_attributesSuccess := THIS^.pLogRecord^.attributes.setStringAttribute(
	key:=key,
	value:=value,
	failureReason=>_attributesFailureReason
);
IF NOT _attributesSuccess THEN
	THIS^._failed := TRUE;
	CASE _attributesFailureReason OF
		E_AttributesFailureReason.MEMORY_ALLOCATION_FAILURE:
			THIS^._failureReason := E_LoggerFailureReason.MEMORY_ALLOCATION_FAILURE;
		E_AttributesFailureReason.ATTRIBUTE_COUNT_LIMIT_REACHED:
			THIS^._failureReason := E_LoggerFailureReason.ATTRIBUTE_COUNT_LIMIT_REACHED;
		E_AttributesFailureReason.KV_VALUE_TYPE_UNSUPPORTED:
			THIS^._failureReason := E_LoggerFailureReason.ATTRIBUTE_VALUE_TYPE_UNSUPPORTED;
	ELSE
		THIS^._failureReason := E_LoggerFailureReason.ATTRIBUTE_VALUE_INVALID;
	END_CASE
END_IF
END_METHOD

METHOD setTimestamp: REFERENCE TO FB_Logger
VAR_INPUT
	timestamp: ULINT;
END_VAR
setTimestamp REF= THIS^;

IF THIS^._shouldReturnEarly() THEN
	RETURN;
END_IF

// if everything above worked, assign the value
THIS^.pLogRecord^.timestamp := timestamp;
END_METHOD

(* Sets the record's trace id from raw bytes. Application code uses setTraceContextFromSpan; this setter is for tests and for setTraceContextFromSpan itself. *)
METHOD _setTraceId: REFERENCE TO FB_Logger
VAR_INPUT
	pBytes: POINTER TO BYTE;
	nSize: UDINT;
END_VAR
VAR
	_pDest: POINTER TO FB_TraceId;
	_factoryFailureReason: E_ValueFactoryFailureReason;
END_VAR
_setTraceId REF= THIS^;

IF THIS^._shouldReturnEarly() THEN
	RETURN;
END_IF

// create an instance of FB_TraceId
IF NOT ValueFactory.createTraceId(
	pDest:=_pDest,
	pBytes:=pBytes,
	nSize:=nSize,
	failureReason=>_factoryFailureReason
	) THEN
	THIS^._failed := TRUE;
	CASE _factoryFailureReason OF
		E_ValueFactoryFailureReason.MEMORY_ALLOCATION_FAILURE:
			THIS^._failureReason := E_LoggerFailureReason.MEMORY_ALLOCATION_FAILURE;
		E_ValueFactoryFailureReason.TRACE_ID_BYTES_POINTER_NULL:
			THIS^._failureReason := E_LoggerFailureReason.TRACE_ID_BYTES_POINTER_NULL;
		E_ValueFactoryFailureReason.TRACE_ID_BYTE_COUNT_TOO_SMALL:
			THIS^._failureReason := E_LoggerFailureReason.TRACE_ID_BYTE_COUNT_TOO_SMALL;
	ELSE
		THIS^._failureReason := E_LoggerFailureReason.TRACE_ID_INVALID;
	END_CASE
	RETURN;
END_IF

// assign to the log record
// delete trace id if it's already set.
IF THIS^.pLogRecord^.traceId <> 0 THEN
	THIS^.pLogRecord^.traceId^.delete(pSelf:=THIS^.pLogRecord^.traceId);
END_IF
// transfer ownership of the data
THIS^.pLogRecord^.traceId := _pDest;
_pDest := 0;
END_METHOD

(*
	This method starts the build process with the required log record state.
	Use the fluent setter methods for optional fields.
	
	Example:
	IF NOT logger
		.startLogRecord(severityNumber := E_SeverityNumber.WARN)
		.setBody('process cycle amps warning, motor fault imminent')
		.setTraceContextFromSpan(pSpan)  // a no-op when pSpan is 0
		.setNumberAttribute('motor.amps.min', minAmps)
		.setNumberAttribute('motor.amps.max', maxAmps)
		.setNumberAttribute('motor.amps.avg', avgAmps)
		.emit(failureResult=>failureResult) THEN
		// CASE failureResult OF ...
	END_IF
*)
METHOD startLogRecord: REFERENCE TO FB_Logger
VAR_INPUT
	severityNumber: E_SeverityNumber;
END_VAR
VAR
	_timestamp: ULINT;
END_VAR
VAR CONSTANT
	UNIX_EPOCH_DIFF: ULINT := 116444736000000000;
END_VAR
startLogRecord REF= THIS^;

// do not replace the first failure in an active fluent chain
IF THIS^.pLogRecord <> 0 THEN
	IF NOT THIS^._failed THEN
		THIS^._failed := TRUE;
		THIS^._failureReason := E_LoggerFailureReason.LOG_RECORD_ALREADY_STARTED;
	END_IF
	RETURN;
END_IF

THIS^._failed := FALSE;
THIS^._failureReason := E_LoggerFailureReason.NA;


_timestamp := (F_GetSystemTime() - UNIX_EPOCH_DIFF) * 100;  // NT ticks (100ns) -> unix epoch nanos


// instantiate a log record
IF NOT THIS^._createLogRecord(
	pDest:=THIS^.pLogRecord,
	severityNumber:=severityNumber,
	timestamp:=_timestamp,
	failureReason=>THIS^._failureReason
	) THEN
	THIS^._failed := TRUE;
END_IF
END_METHOD

END_FUNCTION_BLOCK

// ---- OTEL/LOGGING/PROVIDER/FUNCTION_BLOCKS/FB_LoggerProvider.TcPOU
FUNCTION_BLOCK FB_LoggerProvider
VAR
	_resource: REFERENCE TO FB_Resource; // borrowed; the declaring scope owns its lifetime
	_records: FB_LogRecordQueue(TcOtlp_GVL.MAX_LOG_RECORDS_PER_SCAN);
	_head: POINTER TO ST_LinkedListNode;
	_failureReason: E_LoggerProviderFailureReason;
END_VAR
VAR_OUTPUT
	stagedProcessorCount: UDINT;
END_VAR

METHOD _freeProcessors
VAR
	_idx: UDINT;
	_node: POINTER TO ST_LinkedListNode;
END_VAR
FOR _idx := 0 TO TcOtlp_GVL.MAX_LOOP_COUNT DO
	IF THIS^._head = 0 THEN
		EXIT;
	END_IF
	_node := THIS^._head^.nxt;
	__DELETE(THIS^._head);
	THIS^._head := _node;
	// count down per node, so the count never claims nodes that are gone or hides ones that remain
	IF THIS^.stagedProcessorCount > 0 THEN
		THIS^.stagedProcessorCount := THIS^.stagedProcessorCount - 1;
	END_IF
END_FOR
END_METHOD

//FB_Exit must be implemented explicitly. If there is an implementation, then the
//method is called before the controller removes the code of the function block instance
//(implicit call). The return value is not evaluated.
METHOD FB_Exit: BOOL
VAR_INPUT
    bInCopyCode: BOOL;  // TRUE: the exit method is called in order to leave the instance which will be copied afterwards (online change).  
END_VAR
IF NOT bInCopyCode THEN
	THIS^._freeProcessors();
	THIS^._records.free();
END_IF
END_METHOD

//FB_Init is always available implicitly and it is used primarily for initialization.
//The return value is not evaluated. For a specific influence, you can also declare the
//methods explicitly and provide additional code there with the standard initialization
//code. You can evaluate the return value.
METHOD FB_Init: BOOL
VAR_INPUT
    bInitRetains: BOOL; // TRUE: the retain variables are initialized (reset warm / reset cold)
    bInCopyCode: BOOL;  // TRUE: the instance will be copied to the copy code afterward (online change)
	resource: REFERENCE TO FB_Resource;
END_VAR
THIS^._resource REF= resource;
END_METHOD

METHOD onEmit : BOOL
VAR_IN_OUT
	record: POINTER TO FB_LogRecord;
END_VAR
VAR
	_pushFailureReason: E_LogRecordQueueFailureReason;
END_VAR
onEmit := FALSE;

IF record = 0 THEN
	RETURN;
END_IF

IF NOT THIS^._records.push(pValue:=record, failureReason=>_pushFailureReason) THEN
	RETURN;
END_IF

onEmit := TRUE;
END_METHOD

PROPERTY resource : REFERENCE TO FB_Resource
GET
resource REF= THIS^._resource;
END_GET
END_PROPERTY

METHOD stageProcessor : REFERENCE TO FB_LoggerProvider
VAR_INPUT
	processor: REFERENCE TO FB_LogRecordProcessor_Base;
END_VAR
VAR
	_idx: UDINT;
	_node: POINTER TO ST_LinkedListNode;
END_VAR
stageProcessor REF= THIS^;

// special case if no processors have been registered
IF THIS^._head = 0 THEN
	THIS^._head := __NEW(ST_LinkedListNode);
	IF THIS^._head = 0 THEN
		THIS^._failureReason := E_LoggerProviderFailureReason.STAGE_PROCESSOR_FAILURE;
		RETURN;
	END_IF
	THIS^._head^.val := processor.pSelf;
	THIS^.stagedProcessorCount := THIS^.stagedProcessorCount + 1;
// generic case if at least on processor has been registerd
ELSE
	_node := THIS^._head;
	FOR _idx := 0 TO TcOtlp_GVL.MAX_LOOP_COUNT DO
		IF _node^.val = processor.pSelf THEN
			// silently do nothing if processor already added for this tick
			RETURN;
		ELSIF _node^.nxt = 0 THEN
			// at most MAX_LOOP_COUNT nodes, so _freeProcessors always releases them all
			IF THIS^.stagedProcessorCount >= TcOtlp_GVL.MAX_LOOP_COUNT THEN
				THIS^._failureReason := E_LoggerProviderFailureReason.STAGE_PROCESSOR_FAILURE;
				RETURN;
			END_IF
			_node^.nxt := __NEW(ST_LinkedListNode);
			IF _node^.nxt = 0 THEN
				THIS^._failureReason := E_LoggerProviderFailureReason.STAGE_PROCESSOR_FAILURE;
				RETURN;
			END_IF
			_node^.nxt^.val := processor.pSelf;
			THIS^.stagedProcessorCount := THIS^.stagedProcessorCount + 1;
			RETURN;
		END_IF
		_node := _node^.nxt;
	END_FOR
END_IF
END_METHOD

METHOD tick : BOOL
VAR_OUTPUT
	failureReason: E_LoggerProviderFailureReason;
END_VAR
VAR
	_i: UDINT;
	_j: UDINT;
	_ownedRecordCount: UDINT;
	_node: POINTER TO ST_LinkedListNode;
	_processor: POINTER TO FB_LogRecordProcessor_Base;
	_record: POINTER TO FB_LogRecord;
END_VAR
tick := FALSE;
failureReason := THIS^._failureReason;

// short circuit if fluent calls to add processors failed
IF failureReason <> E_LoggerProviderFailureReason.NA THEN
	RETURN;
END_IF

// if no processors added skip loop iteration and just free the queue
IF THIS^._head = 0 THEN
	THIS^._records.free();
	tick := TRUE;
	RETURN;
END_IF

// loop over each item and call each processor for each record
_ownedRecordCount := THIS^._records.count;
FOR _i := 1 TO _ownedRecordCount DO
	IF NOT THIS^._records.pop(_record) THEN
		failureReason := E_LoggerProviderFailureReason.QUEUE_POP_FAILURE;
		JMP _endLabel;
	END_IF
	// call on emit for each record
	_node := THIS^._head;
	FOR _j := 1 TO THIS^.stagedProcessorCount DO
		IF _node = 0 THEN
			failureReason := E_LoggerProviderFailureReason.UNEXPECTED_NULL_LINKED_LIST_NODE;
			JMP _endLabel;
		END_IF
		_processor := _node^.val;
		IF _processor = 0 THEN
			failureReason := E_LoggerProviderFailureReason.UNEXPECTED_NULL_PROCESSOR_POINTER;
			JMP _endLabel;
		END_IF
		_processor^.onEmit(_record^);
		_node := _node^.nxt;
	END_FOR
	_record^.delete(pSelf:=_record);
END_FOR

// tick each processor
_node := THIS^._head;
FOR _j := 1 TO THIS^.stagedProcessorCount DO
	// guard before dereferencing; walking off the tail on the last iteration is
	// normal termination, so only a list shorter than the count is a failure
	IF _node = 0 THEN
		failureReason := E_LoggerProviderFailureReason.UNEXPECTED_NULL_LINKED_LIST_NODE;
		JMP _endLabel;
	END_IF
	_processor := _node^.val;
	IF _processor = 0 THEN
		failureReason := E_LoggerProviderFailureReason.UNEXPECTED_NULL_PROCESSOR_POINTER;
		JMP _endLabel;
	END_IF
	_processor^.tick();
	_node := _node^.nxt;
END_FOR

// clean up and return
_endLabel:
THIS^._records.free();
THIS^._freeProcessors();
IF _record <> 0 THEN _record^.delete(pSelf:=_record); END_IF
tick := failureReason = E_LoggerProviderFailureReason.NA;
END_METHOD

END_FUNCTION_BLOCK

// ---- OTEL/LOGGING/PROCESSORS/FUNCTION_BLOCKS/FB_LogRecordProcessor_Base.TcPOU
FUNCTION_BLOCK ABSTRACT FB_LogRecordProcessor_Base

METHOD ABSTRACT enrich
VAR_IN_OUT
	logRecord: FB_LogRecord;
END_VAR
END_METHOD

METHOD ABSTRACT free
VAR_INPUT
END_VAR
END_METHOD

METHOD ABSTRACT onEmit
VAR_INPUT
	logRecord: REFERENCE TO FB_LogRecord;
END_VAR
END_METHOD

PROPERTY pSelf : POINTER TO FB_LogRecordProcessor_Base
GET
pSelf := THIS;
END_GET
END_PROPERTY

METHOD ABSTRACT tick
END_METHOD

END_FUNCTION_BLOCK

// ---- OTEL/LOGGING/PROCESSORS/FUNCTION_BLOCKS/FB_LogRecordProcessor_Batch.TcPOU
(*
	Batch processor. onEmit enriches and stores records only. Call the FB body
	cyclically to advance the exporter and export the oldest queued records when
	the schedule delay elapses or a full batch is available.
*)
FUNCTION_BLOCK FB_LogRecordProcessor_Batch EXTENDS FB_LogRecordProcessor_Base;
VAR_OUTPUT
	scheduledDelayMillis: UDINT := 1000;	// maximum delay before queued records are exported
	maxExportBatchSize: UDINT := 512;		// maximum records transferred to one export
	lastOperationSucceeded: BOOL := TRUE;
	failureResult: E_LogRecordProcessorFailureReason;
END_VAR
VAR
	_scheduleDelayTimer: TON;
	_records: FB_LogRecordQueue(maxCount:=0);  // set again during THIS^.FB_Init
	_exporter: REFERENCE TO FB_LogRecordExporter_Base;
	_rejectedCount: UDINT;  // records that could not be cloned or queued
END_VAR

// no-op; override to change log mutation/enrichment functionality
METHOD enrich
VAR_IN_OUT
	logRecord: FB_LogRecord;
END_VAR
END_METHOD

METHOD exportIfNeeded
VAR
	_exportFailureReason: E_LogRecordExporterFailureReason;
END_VAR
IF THIS^.maxExportBatchSize = 0
	OR_ELSE NOT __ISVALIDREF(THIS^._exporter)
	OR_ELSE THIS^._exporter.isBusy()
	OR_ELSE THIS^._records.count = 0 THEN
	RETURN;
END_IF

IF NOT THIS^._scheduleDelayTimer.Q
	AND_THEN THIS^._records.count < THIS^.maxExportBatchSize THEN
	RETURN;
END_IF

IF THIS^._exporter.export(
	logRecords:=THIS^._records,
	count:=THIS^.maxExportBatchSize,
	failureReason=>_exportFailureReason
) THEN
	THIS^._scheduleDelayTimer(IN:=FALSE, PT:=UDINT_TO_TIME(THIS^.scheduledDelayMillis));
	THIS^.lastOperationSucceeded := TRUE;
	THIS^.failureResult := E_LogRecordProcessorFailureReason.NA;
ELSE
	THIS^.lastOperationSucceeded := FALSE;
	THIS^.failureResult := E_LogRecordProcessorFailureReason.EXPORT_FAILURE;
END_IF
END_METHOD

METHOD FB_Exit : BOOL
VAR_INPUT
	bInCopyCode: BOOL;
END_VAR
IF NOT bInCopyCode THEN
	THIS^.free();
END_IF
END_METHOD

//FB_Init is always available implicitly and it is used primarily for initialization.
//The return value is not evaluated. For a specific influence, you can also declare the
//methods explicitly and provide additional code there with the standard initialization
//code. You can evaluate the return value.
METHOD FB_Init: BOOL
VAR_INPUT
    bInitRetains: BOOL; // TRUE: the retain variables are initialized (reset warm / reset cold)
    bInCopyCode: BOOL;  // TRUE: the instance will be copied to the copy code afterward (online change)
	maxQueueSize: UDINT := 2048;			// zero is unbounded; otherwise the oldest record is dropped when full
	scheduledDelayMillis: UDINT := 1000;	// maximum delay before queued records are exported
	maxExportBatchSize: UDINT := 512;		// maximum records transferred to one export
	exporter: REFERENCE TO FB_LogRecordExporter_Base;	// the exporter where the LogRecords are pushed.
END_VAR
THIS^._records.FB_Init(FALSE, FALSE, maxQueueSize);
THIS^.scheduledDelayMillis := scheduledDelayMillis;
THIS^.maxExportBatchSize := maxExportBatchSize;
IF __ISVALIDREF(exporter) THEN
	THIS^._exporter REF= exporter;
END_IF
END_METHOD

METHOD free
THIS^._records.free();
THIS^._scheduleDelayTimer(IN:=FALSE, PT:=UDINT_TO_TIME(THIS^.scheduledDelayMillis));
END_METHOD

(*
	Clones the log record onto the tail of the arrival-order queue.
	When the queue holds maxQueueSize records, the oldest record is
	dropped from the head to make room for the newest.
*)
METHOD onEmit
VAR_INPUT
	logRecord: REFERENCE TO FB_LogRecord;
END_VAR
VAR
	_pRecord: POINTER TO FB_LogRecord;
	_cloneFailureResult: E_LogRecordCloneFailureReason;
	_queueFailureReason: E_LogRecordQueueFailureReason;
END_VAR
THIS^.enrich(logRecord);

IF __ISVALIDREF(THIS^._exporter) THEN
	_pRecord := 0;
	IF NOT logRecord.cloneTo(pDest:=_pRecord, failureReason=>_cloneFailureResult) THEN
		IF _pRecord <> 0 THEN _pRecord^.delete(pSelf:=_pRecord); END_IF
		THIS^._rejectedCount := THIS^._rejectedCount + 1;
		THIS^.lastOperationSucceeded := FALSE;
		THIS^.failureResult := E_LogRecordProcessorFailureReason.RECORD_CLONE_FAILURE;
		RETURN;
	END_IF
	
	IF NOT THIS^._records.push(pValue:=_pRecord, failureReason=>_queueFailureReason) THEN
		_pRecord^.delete(pSelf:=_pRecord);
		THIS^._rejectedCount := THIS^._rejectedCount + 1;
		THIS^.lastOperationSucceeded := FALSE;
		THIS^.failureResult := E_LogRecordProcessorFailureReason.QUEUE_PUSH_FAILURE;
		RETURN;
	END_IF
END_IF

THIS^.lastOperationSucceeded := TRUE;
THIS^.failureResult := E_LogRecordProcessorFailureReason.NA;
END_METHOD

METHOD tick
VAR
	_exportFailureReason: E_LogRecordExporterFailureReason;
END_VAR
THIS^._scheduleDelayTimer(
	IN:=THIS^._records.count > 0,
	PT:=UDINT_TO_TIME(THIS^.scheduledDelayMillis)
);

IF __ISVALIDREF(THIS^._exporter) THEN
	THIS^._exporter.tick(failureReason=>_exportFailureReason);
	THIS^.exportIfNeeded();
END_IF
END_METHOD

(* Records lost so far: evicted from a full queue, or not cloned or queued. *)
PROPERTY droppedCount : UDINT
GET
droppedCount := THIS^._records.droppedCount + THIS^._rejectedCount;
END_GET
END_PROPERTY

(* Records waiting for export. *)
PROPERTY queuedCount : UDINT
GET
queuedCount := THIS^._records.count;
END_GET
END_PROPERTY

END_FUNCTION_BLOCK

// ---- OTEL/LOGGING/PROCESSORS/FUNCTION_BLOCKS/FB_LogRecordProcessor_Simple.TcPOU
FUNCTION_BLOCK FB_LogRecordProcessor_Simple EXTENDS FB_LogRecordProcessor_Base;
VAR
	_records: FB_LogRecordQueue(maxCount:=1);
	_exporter: REFERENCE TO FB_LogRecordExporter_Base;
END_VAR

// no-op, overwride to change log mutation/enrichment functionality
METHOD enrich
VAR_IN_OUT
	logRecord	: FB_LogRecord;
END_VAR
END_METHOD

//FB_Exit must be implemented explicitly. If there is an implementation, then the
//method is called before the controller removes the code of the function block instance
//(implicit call). The return value is not evaluated.
METHOD FB_Exit: BOOL
VAR_INPUT
    bInCopyCode: BOOL;  // TRUE: the exit method is called in order to leave the instance which will be copied afterwards (online change).  
END_VAR
IF NOT bInCopyCode THEN
	THIS^.free();
END_IF
END_METHOD

//FB_Init is always available implicitly and it is used primarily for initialization.
//The return value is not evaluated. For a specific influence, you can also declare the
//methods explicitly and provide additional code there with the standard initialization
//code. You can evaluate the return value.
METHOD FB_Init: BOOL
VAR_INPUT
    bInitRetains: BOOL; // TRUE: the retain variables are initialized (reset warm / reset cold)
    bInCopyCode: BOOL;  // TRUE: the instance will be copied to the copy code afterward (online change)
	exporter: REFERENCE TO FB_LogRecordExporter_Base;
END_VAR
IF __ISVALIDREF(exporter) THEN
	THIS^._exporter REF= exporter;
ELSE
	THIS^._exporter REF= 0;
END_IF
END_METHOD

METHOD free
THIS^._records.free();
END_METHOD

METHOD onEmit
VAR_INPUT
	logRecord: REFERENCE TO FB_LogRecord;
END_VAR
VAR
	_pLogRecord: POINTER TO FB_LogRecord;
	_cloneFailureResult: E_LogRecordCloneFailureReason;
	_queueFailureReason: E_LogRecordQueueFailureReason;
	_exportFailureReason: E_LogRecordExporterFailureReason;
END_VAR
THIS^.enrich(logRecord);

IF __ISVALIDREF(THIS^._exporter) THEN
	IF (NOT THIS^._exporter.isBusy()) THEN
		IF logRecord.cloneTo(pDest:=_pLogRecord, failureReason=>_cloneFailureResult) THEN
			IF THIS^._records.push(pValue:=_pLogRecord, failureReason=>_queueFailureReason) THEN
				THIS^._exporter.export(
					logRecords:=THIS^._records,
					count:=1,
					failureReason=>_exportFailureReason
				);
			END_IF
		END_IF
	END_IF
END_IF

// If the exporter did not accept the buffer, the simple processor drops it.
THIS^.free();
IF _pLogRecord <> 0 THEN _pLogRecord^.delete(pSelf:=_pLogRecord); END_IF
END_METHOD

METHOD tick
VAR
	_exportFailureReason: E_LogRecordExporterFailureReason;
END_VAR
IF __ISVALIDREF(THIS^._exporter) THEN
	THIS^._exporter.tick(failureReason=>_exportFailureReason);
END_IF
END_METHOD

END_FUNCTION_BLOCK

// ---- OTEL/TRACING/EXPORTING/FUNCTION_BLOCKS/FB_SpanExporter_Base.TcPOU
(*
	Contract shared by span exporters. A processor offers a batch with export, which moves up to
	count of the oldest spans out of the processor's queue into the exporter without cloning
	them. The exporter owns the batch until free, which runs when the batch is delivered or
	failed, when the next batch is accepted, and when the exporter is destroyed.
	Concrete exporters advance delivery in tick and report through isBusy whether they can take
	another batch. Only ended spans reach an exporter.
*)
FUNCTION_BLOCK ABSTRACT FB_SpanExporter_Base
VAR
	_spans: FB_SpanQueue(maxCount:=0);
	_exportActive: BOOL;
	_callFailureReason: E_SpanExporterFailureReason;
END_VAR

(*
	Takes ownership of up to count of the oldest spans in spans. While busy it refuses with
	ACTIVE_EXPORT_IN_PROGRESS and leaves spans unchanged. A count of zero accepts nothing and
	succeeds.
*)
METHOD export : BOOL
VAR_IN_OUT
	spans: FB_SpanQueue;  // accepted spans are transferred out of this queue
END_VAR
VAR_INPUT
	count: UDINT;
END_VAR
VAR_OUTPUT
	failureReason: E_SpanExporterFailureReason;
END_VAR
VAR
	_queueFailureReason: E_SpanQueueFailureReason;
END_VAR
export := FALSE;
failureReason := E_SpanExporterFailureReason.NA;

IF THIS^.isBusy() THEN
	failureReason := E_SpanExporterFailureReason.ACTIVE_EXPORT_IN_PROGRESS;
	RETURN;
END_IF

// release a finished batch still held by the exporter before accepting the next one
THIS^.free();
IF NOT spans.transferTo(
	destination:=THIS^._spans,
	count:=count,
	failureReason=>_queueFailureReason
) THEN
	failureReason := E_SpanExporterFailureReason.QUEUE_TRANSFER_FAILURE;
	RETURN;
END_IF

THIS^._exportActive := THIS^._spans.count > 0;
export := TRUE;
END_METHOD

METHOD FB_Exit : BOOL
VAR_INPUT
	bInCopyCode: BOOL;
END_VAR
IF NOT bInCopyCode THEN
	THIS^.free();
END_IF
END_METHOD

(* Releases every span the exporter owns and clears the active export. *)
METHOD free
THIS^._spans.free();
THIS^._exportActive := FALSE;
END_METHOD

(* TRUE while the exporter cannot accept another batch. *)
METHOD ABSTRACT isBusy : BOOL
END_METHOD

(* Advances delivery of the accepted batch. Call it every scan. *)
METHOD ABSTRACT tick : BOOL
VAR_OUTPUT
	failureReason: E_SpanExporterFailureReason;
END_VAR
END_METHOD

END_FUNCTION_BLOCK

// ---- OTEL/TRACING/SPAN/FUNCTION_BLOCKS/FB_SpanQueue.TcPOU
(*
	FIFO queue that owns every FB_Span pointer it contains. push takes ownership and
	clears the caller's pointer; pop hands ownership back. push drops the oldest owned
	spans when the bound is reached. The bound is maxCount, but never more than
	TcOtlp_GVL.MAX_LOOP_COUNT: a maxCount of zero, or one above that limit, is held to
	MAX_LOOP_COUNT so that free always reaches the end.
	reset and next walk the spans oldest first without taking ownership. rotate moves the
	oldest span to the back, so a consumer can skip it and keep arrival order. transferTo moves the oldest spans into another queue, for handing
	a batch to an exporter.
*)
FUNCTION_BLOCK FB_SpanQueue
VAR
	_head: POINTER TO ST_LinkedListNode;
	_tail: POINTER TO ST_LinkedListNode;
	_cursor: POINTER TO ST_LinkedListNode;  // next node returned by next; 0 at the end
END_VAR
VAR_OUTPUT
	count: UDINT;
	maxCount: UDINT;
	droppedCount: UDINT;
END_VAR

(* The enforced bound: maxCount, held to MAX_LOOP_COUNT when it is zero or larger. *)
METHOD _capacity : UDINT
IF THIS^.maxCount = 0 OR THIS^.maxCount > TcOtlp_GVL.MAX_LOOP_COUNT THEN
	_capacity := TcOtlp_GVL.MAX_LOOP_COUNT;
ELSE
	_capacity := THIS^.maxCount;
END_IF
END_METHOD

METHOD FB_Exit : BOOL
VAR_INPUT
	bInCopyCode: BOOL;
END_VAR
IF NOT bInCopyCode THEN
	THIS^.free();
END_IF
END_METHOD

METHOD FB_Init : BOOL
VAR_INPUT
	bInitRetains: BOOL;
	bInCopyCode: BOOL;
	maxCount: UDINT := 0;
END_VAR
THIS^.maxCount := maxCount;
END_METHOD

(*
	Releases every owned span. push holds count to MAX_LOOP_COUNT, so the loop always
	reaches the end. If it ever stops early, the unreleased nodes stay in the queue and
	free returns FALSE, so a later call can finish the job.
*)
METHOD free : BOOL
VAR
	_idx: UDINT;
	_node: POINTER TO ST_LinkedListNode;
	_span: POINTER TO FB_Span;
END_VAR
FOR _idx := 0 TO TcOtlp_GVL.MAX_LOOP_COUNT DO
	IF THIS^._head = 0 THEN
		EXIT;
	END_IF

	_node := THIS^._head;
	THIS^._head := _node^.nxt;
	IF _node^.val <> 0 THEN
		_span := _node^.val;
		_node^.val := 0;
		_span^.delete(pSelf:=_span);
	END_IF
	__DELETE(_node);
	_node := 0;
	IF THIS^.count > 0 THEN
		THIS^.count := THIS^.count - 1;
	END_IF
END_FOR

IF THIS^._head = 0 THEN
	THIS^._tail := 0;
	THIS^.count := 0;
END_IF
THIS^._cursor := THIS^._head;
free := THIS^._head = 0;
END_METHOD

(*
	Returns the span at the cursor and advances it, or 0 after the last span. The span is
	borrowed: the queue still owns it, and it is valid only until it is popped or dropped.
	Call reset first.
*)
METHOD next : POINTER TO FB_Span
next := 0;
IF THIS^._cursor <> 0 THEN
	next := THIS^._cursor^.val;
	THIS^._cursor := THIS^._cursor^.nxt;
END_IF
END_METHOD

(* Moves the oldest span to pValue, which must be 0. The caller owns it on success. *)
METHOD pop : BOOL
VAR_IN_OUT
	pValue: POINTER TO FB_Span;
END_VAR
VAR_OUTPUT
	failureReason: E_SpanQueueFailureReason;
END_VAR
VAR
	_node: POINTER TO ST_LinkedListNode;
END_VAR
pop := FALSE;
failureReason := E_SpanQueueFailureReason.NA;

IF pValue <> 0 THEN
	failureReason := E_SpanQueueFailureReason.DESTINATION_ALREADY_ASSIGNED;
	RETURN;
END_IF
IF THIS^._head = 0 THEN
	failureReason := E_SpanQueueFailureReason.QUEUE_EMPTY;
	RETURN;
END_IF

_node := THIS^._head;
THIS^._head := _node^.nxt;
IF THIS^._head = 0 THEN
	THIS^._tail := 0;
END_IF
IF THIS^._cursor = _node THEN
	THIS^._cursor := THIS^._head;
END_IF

pValue := _node^.val;
_node^.val := 0;
_node^.nxt := 0;
__DELETE(_node);
_node := 0;
THIS^.count := THIS^.count - 1;
pop := failureReason = E_SpanQueueFailureReason.NA;
END_METHOD

(*
	Takes ownership of the span and clears pValue. On failure pValue is left unchanged
	and still owned by the caller.
*)
METHOD push : BOOL
VAR_IN_OUT
	pValue: POINTER TO FB_Span;
END_VAR
VAR_OUTPUT
	failureReason: E_SpanQueueFailureReason;
END_VAR
VAR
	_node: POINTER TO ST_LinkedListNode;
	_droppedSpan: POINTER TO FB_Span;
	_popFailureReason: E_SpanQueueFailureReason;
	_idx: UDINT;
	_bound: UDINT;
END_VAR
push := FALSE;
failureReason := E_SpanQueueFailureReason.NA;

IF pValue = 0 THEN
	failureReason := E_SpanQueueFailureReason.SPAN_POINTER_NULL;
	RETURN;
END_IF

// Allocate before evicting so an allocation failure leaves the queue unchanged.
_node := __NEW(ST_LinkedListNode);
IF _node = 0 THEN
	failureReason := E_SpanQueueFailureReason.MEMORY_ALLOCATION_FAILURE;
	RETURN;
END_IF

// maxCount is writable, so also restore the bound after a runtime reduction.
_bound := THIS^._capacity();
FOR _idx := 0 TO TcOtlp_GVL.MAX_LOOP_COUNT DO
	IF THIS^.count < _bound THEN
		EXIT;
	END_IF
	IF NOT THIS^.pop(pValue:=_droppedSpan, failureReason=>_popFailureReason) THEN
		__DELETE(_node);
		_node := 0;
		failureReason := _popFailureReason;
		RETURN;
	END_IF
	_droppedSpan^.delete(pSelf:=_droppedSpan);
	THIS^.droppedCount := THIS^.droppedCount + 1;
END_FOR
IF THIS^.count >= _bound THEN
	__DELETE(_node);
	_node := 0;
	failureReason := E_SpanQueueFailureReason.MAX_SIZE_ENFORCEMENT_FAILURE;
	RETURN;
END_IF

_node^.val := pValue;
_node^.nxt := 0;
IF THIS^._tail = 0 THEN
	THIS^._head := _node;
ELSE
	THIS^._tail^.nxt := _node;
END_IF
THIS^._tail := _node;
THIS^.count := THIS^.count + 1;
pValue := 0;
push := failureReason = E_SpanQueueFailureReason.NA;
END_METHOD

(* Moves the cursor to the oldest span, so next starts from the head. *)
METHOD reset
THIS^._cursor := THIS^._head;
END_METHOD

(*
	Moves up to count of the oldest spans into destination, which must be empty. Ownership moves
	with the nodes, so nothing is cloned or released. The move stops at this queue's count and at
	the destination's bound.
*)
METHOD transferTo : BOOL
VAR_IN_OUT
	destination: FB_SpanQueue;
END_VAR
VAR_INPUT
	count: UDINT;
END_VAR
VAR_OUTPUT
	failureReason: E_SpanQueueFailureReason;
END_VAR
VAR
	_transferCount: UDINT;
	_idx: UDINT;
END_VAR
transferTo := FALSE;
failureReason := E_SpanQueueFailureReason.NA;

IF ADR(destination) = THIS THEN
	failureReason := E_SpanQueueFailureReason.SELF_TRANSFER_NOT_ALLOWED;
	RETURN;
END_IF
IF destination.count <> 0 OR_ELSE destination._head <> 0 OR_ELSE destination._tail <> 0 THEN
	failureReason := E_SpanQueueFailureReason.DESTINATION_NOT_EMPTY;
	RETURN;
END_IF

_transferCount := MIN(count, THIS^.count, destination._capacity());
IF _transferCount = 0 THEN
	transferTo := TRUE;
	RETURN;
END_IF

// count never exceeds MAX_LOOP_COUNT, so this walk is bounded
destination._head := THIS^._head;
destination._tail := destination._head;
FOR _idx := 1 TO _transferCount - 1 DO
	destination._tail := destination._tail^.nxt;
END_FOR

THIS^._head := destination._tail^.nxt;
destination._tail^.nxt := 0;
destination._cursor := destination._head;
destination.count := _transferCount;

THIS^.count := THIS^.count - _transferCount;
THIS^._cursor := THIS^._head;
IF THIS^._head = 0 THEN
	THIS^._tail := 0;
END_IF
transferTo := TRUE;
END_METHOD

(* Moves the oldest span to the back without changing ownership, and resets the cursor. *)
METHOD rotate : BOOL
VAR_OUTPUT
	failureReason: E_SpanQueueFailureReason;
END_VAR
VAR
	_node: POINTER TO ST_LinkedListNode;
END_VAR
rotate := FALSE;
failureReason := E_SpanQueueFailureReason.NA;

IF THIS^._head = 0 THEN
	failureReason := E_SpanQueueFailureReason.QUEUE_EMPTY;
	RETURN;
END_IF

IF THIS^._head <> THIS^._tail THEN
	_node := THIS^._head;
	THIS^._head := _node^.nxt;
	_node^.nxt := 0;
	THIS^._tail^.nxt := _node;
	THIS^._tail := _node;
END_IF

THIS^._cursor := THIS^._head;
rotate := failureReason = E_SpanQueueFailureReason.NA;
END_METHOD

END_FUNCTION_BLOCK

// ---- OTEL/TRACING/EXPORTING/FUNCTION_BLOCKS/FB_SpanExporter_File.TcPOU
(*
	Appends each accepted batch to a file as one OTLP ProtoJSON TracesData object per line
	(JSON Lines), grouped by resource and scope. The file is opened in append mode and closed
	again for every batch. Call the instance, or tick, every scan: the exporter is busy from
	export until currentState reaches done or error. The batch is released at either end, and
	an error is reported by tick until the next batch is accepted.
*)
FUNCTION_BLOCK FB_SpanExporter_File EXTENDS FB_SpanExporter_Base
VAR_OUTPUT
	currentState: E_FileExporterState;
END_VAR
VAR
	_execute: BOOL;
	_filepath: T_MaxString;
	_hFile: UINT;
	_len: UDINT;
	_execRTrig: R_TRIG;
	_pString: POINTER TO STRING;  // payload buffer, owned while a write is in flight
	_jsonVal: SJsonValue;
	_resourceSpansArray: SJsonValue;
	_fileOpener: FB_FileOpen;
	_fileWriter: FB_FileWrite;
	_fileCloser: FB_FileClose;
	_computedState: E_FileExporterState;
	_failureReason: E_SpanExporterFailureReason;
	_serializationFailureReason: E_ProtoJsonSerializerFailureReason;
	_serializer: FB_SpanProtoJsonSerializer;
END_VAR

THIS^.tick(failureReason=>THIS^._callFailureReason);

METHOD export : BOOL
VAR_IN_OUT
	spans: FB_SpanQueue;
END_VAR
VAR_INPUT
	count: UDINT;
END_VAR
VAR_OUTPUT
	failureReason: E_SpanExporterFailureReason;
END_VAR
// a finished exporter accepts the next batch at once
IF THIS^.currentState = E_FileExporterState.done OR THIS^.currentState = E_FileExporterState.error THEN
	THIS^.currentState := E_FileExporterState.idle;
	THIS^._computedState := E_FileExporterState.idle;
END_IF
export := SUPER^.export(
	spans:=spans,
	count:=count,
	failureReason=>failureReason
);
IF export THEN
	THIS^._failureReason := E_SpanExporterFailureReason.NA;
	THIS^._serializationFailureReason := E_ProtoJsonSerializerFailureReason.NA;
END_IF
END_METHOD

(*
	Releases a payload buffer that is still in flight. The FB_FileWrite reading it is
	destroyed with this instance, so nothing uses the buffer afterwards. TwinCAT then
	runs FB_SpanExporter_Base.FB_Exit, which releases the accepted spans.
*)
METHOD FB_Exit : BOOL
VAR_INPUT
	bInCopyCode: BOOL;  // TRUE: the instance is being copied during an online change
END_VAR
// during an online change the copy keeps the buffer, so it must not be released here
IF NOT bInCopyCode AND _pString <> 0 THEN
	__DELETE(_pString);
	_pString := 0;
END_IF
END_METHOD

METHOD FB_Init : BOOL
VAR_INPUT
	bInitRetains: BOOL;  // TRUE: the retain variables are initialized (reset warm / reset cold)
	bInCopyCode: BOOL;  // TRUE: the instance will be copied to the copy code afterward (online change)
	filepath: T_MaxString;  // file the batches are appended to
END_VAR
THIS^._filepath := filepath;
END_METHOD

METHOD isBusy : BOOL
isBusy := THIS^._exportActive;
END_METHOD

METHOD tick : BOOL
VAR_OUTPUT
	failureReason: E_SpanExporterFailureReason;
END_VAR
tick := TRUE;
failureReason := E_SpanExporterFailureReason.NA;

_execute := THIS^._exportActive;
_execRTrig(CLK := _execute AND_THEN THIS^._spans.count > 0);

CASE currentState OF
	E_FileExporterState.idle:
		IF _execRTrig.Q THEN
			_failureReason := E_SpanExporterFailureReason.NA;
			_serializationFailureReason := E_ProtoJsonSerializerFailureReason.NA;
			_computedState := E_FileExporterState.serializing;
		END_IF

	E_FileExporterState.serializing:
		IF NOT _serializer.serializeTracesData(
			spans:=THIS^._spans,
			failureReason=>_serializationFailureReason
		) THEN
			_failureReason := E_SpanExporterFailureReason.SERIALIZATION_FAILURE;
			_computedState := E_FileExporterState.error;
		ELSE
			_jsonVal := _serializer.jsonValue;
			IF _jsonVal = 0 OR_ELSE NOT _serializer.parser.IsObject(_jsonVal) THEN
				_failureReason := E_SpanExporterFailureReason.SERIALIZATION_FAILURE;
				_computedState := E_FileExporterState.error;
			ELSE
				_resourceSpansArray := _serializer.parser.FindMember(_jsonVal, 'resourceSpans');
				IF _resourceSpansArray = 0 OR_ELSE NOT _serializer.parser.IsArray(_resourceSpansArray) THEN
					_failureReason := E_SpanExporterFailureReason.SERIALIZATION_FAILURE;
					_computedState := E_FileExporterState.error;
				ELSE
					_computedState := E_FileExporterState.opening;
				END_IF
			END_IF
		END_IF

	E_FileExporterState.opening:
		IF _fileOpener.bError THEN
			_failureReason := E_SpanExporterFailureReason.FILE_OPEN_FAILURE;
			_computedState := E_FileExporterState.error;
		ELSIF NOT _fileOpener.bBusy THEN
			_hFile := _fileOpener.hFile;
			_computedState := E_FileExporterState.buffering;
		END_IF

	E_FileExporterState.buffering:
		// write one complete TracesData object per JSONL line
		_len := _serializer.parser.GetJsonLength(_jsonVal);  // includes the null terminating character
		IF _len = 0 THEN
			_failureReason := E_SpanExporterFailureReason.SERIALIZATION_FAILURE;
			_computedState := E_FileExporterState.closing;
		ELSE
			_pString := __NEW(BYTE, (_len + 1));  // + 1 for the new line
			IF _pString = 0 THEN
				_failureReason := E_SpanExporterFailureReason.BUFFER_ALLOCATION_FAILURE;
				_computedState := E_FileExporterState.closing;
			ELSE
				_serializer.parser.CopyJson(_jsonVal, _pString^, _len);
				CONCAT2(_pString, ADR('$N'), _pString, _len + 1);
				_computedState := E_FileExporterState.writing;
			END_IF
		END_IF

	E_FileExporterState.writing:
		IF _fileWriter.bError THEN
			IF _pString <> 0 THEN __DELETE(_pString); _pString := 0; END_IF
			_failureReason := E_SpanExporterFailureReason.FILE_WRITE_FAILURE;
			_computedState := E_FileExporterState.closing;
		ELSIF NOT _fileWriter.bBusy THEN
			IF _pString <> 0 THEN __DELETE(_pString); _pString := 0; END_IF
			_computedState := E_FileExporterState.closing;
		END_IF

	E_FileExporterState.closing:
		IF _fileCloser.bError THEN
			IF _failureReason = E_SpanExporterFailureReason.NA THEN
				_failureReason := E_SpanExporterFailureReason.FILE_CLOSE_FAILURE;
			END_IF
			_computedState := E_FileExporterState.error;
		ELSIF NOT _fileCloser.bBusy THEN
			IF _failureReason = E_SpanExporterFailureReason.NA THEN
				_computedState := E_FileExporterState.done;
			ELSE
				_computedState := E_FileExporterState.error;
			END_IF
		END_IF

	E_FileExporterState.done:
		IF NOT _execute THEN
			_computedState := E_FileExporterState.idle;
		END_IF

	E_FileExporterState.error:
		// keep the failure until export accepts a new batch
END_CASE

currentState := _computedState;

IF currentState <= E_FileExporterState.serializing THEN _hFile := 0; END_IF
IF currentState = E_FileExporterState.done
	OR_ELSE currentState = E_FileExporterState.error THEN
	THIS^.free();
END_IF

_fileOpener(
	sNetId:='',
	sPathName:=THIS^._filepath,
	bExecute:=currentState = E_FileExporterState.opening,
	nMode:=FOPEN_MODEAPPEND OR FOPEN_MODETEXT,
	ePath:=PATH_GENERIC,
	tTimeout:=DEFAULT_ADS_TIMEOUT
);

_fileWriter(
	hFile:=_hFile,
	bExecute:=currentState = E_FileExporterState.writing,
	pWriteBuff:=_pString,
	cbWriteLen:=_len
);

_fileCloser(
	hFile:=_hFile,
	bExecute:=currentState = E_FileExporterState.closing
);

IF currentState = E_FileExporterState.error THEN
	tick := FALSE;
	failureReason := _failureReason;
END_IF
END_METHOD

END_FUNCTION_BLOCK

// ---- OTEL/TRACING/SERIALIZATION/FUNCTION_BLOCKS/FB_SpanProtoJsonSerializer.TcPOU
(*
	Writes ended spans as OTLP ProtoJSON: TracesData > ResourceSpans > ScopeSpans > Span.
	serializeTracesData takes ownership of the queued spans and drains the queue: every span
	is released once written, and whatever is left is released on failure.

	Example:
	IF serializer.serializeTracesData(spans:=queue, failureReason=>reason) THEN
		// serializer.parser and serializer.jsonValue hold the document
	END_IF
*)
FUNCTION_BLOCK FB_SpanProtoJsonSerializer EXTENDS FB_BaseProtoJsonSerializer

(*
	Writes the span's links as a 'links' array of Link objects, in the order they were added.
	Walking the links moves their cursor, but the links themselves are only read.
*)
METHOD _serializeLinks : BOOL
VAR_IN_OUT
	v: SJsonValue;
	links: FB_Links;
END_VAR
VAR_OUTPUT
	failureReason: E_ProtoJsonSerializerFailureReason;
END_VAR
VAR
	_array: SJsonValue;
	_obj: SJsonValue;
	_pLink: POINTER TO FB_Link;
	_idx: UDINT;
END_VAR
_serializeLinks := FALSE;
failureReason := E_ProtoJsonSerializerFailureReason.NA;
IF v = 0 THEN
	failureReason := E_ProtoJsonSerializerFailureReason.JSON_VALUE_INVALID;
	RETURN;
END_IF

_array := THIS^.parser.AddArrayMember(v, 'links', 0);
IF _array = 0 THEN
	failureReason := E_ProtoJsonSerializerFailureReason.JSON_OPERATION_FAILURE;
	RETURN;
END_IF

links.reset();
FOR _idx := 0 TO TcOtlp_GVL.MAX_LOOP_COUNT DO
	_pLink := links.next();
	IF _pLink = 0 THEN
		_serializeLinks := TRUE;
		RETURN;
	END_IF

	_obj := THIS^.parser.PushbackJsonValue(_array, '{}');
	IF _obj = 0 THEN
		failureReason := E_ProtoJsonSerializerFailureReason.JSON_OPERATION_FAILURE;
		RETURN;
	END_IF
	IF _pLink^.traceId <> 0 AND_THEN NOT THIS^.serializeTraceIdValue(_obj, _pLink^.traceId, failureReason=>failureReason) THEN RETURN; END_IF
	IF _pLink^.spanId <> 0 AND_THEN NOT THIS^.serializeSpanIdValue(_obj, _pLink^.spanId, failureReason=>failureReason) THEN RETURN; END_IF
	IF _pLink^.traceState <> 0 AND_THEN NOT THIS^._serializeTraceState(_obj, _pLink^.traceState, failureReason=>failureReason) THEN RETURN; END_IF
	IF _pLink^.attributes.count > 0 AND_THEN NOT THIS^.serializeKeyValues(_obj, ADR('attributes'), ADR(_pLink^.attributes), failureReason=>failureReason) THEN RETURN; END_IF
	IF _pLink^.attributes.droppedCount > 0 AND_THEN NOT THIS^.serializeUint32Value(
		_obj,
		ADR('droppedAttributesCount'),
		_pLink^.attributes.droppedCount,
		failureReason=>failureReason
	) THEN
		RETURN;
	END_IF
	IF _pLink^.flags <> 0 AND_THEN NOT THIS^.serializeUint32Value(_obj, ADR('flags'), _pLink^.flags, failureReason=>failureReason) THEN RETURN; END_IF
END_FOR

// FB_Links holds at most MAX_LOOP_COUNT links, so the walk always ends above
failureReason := E_ProtoJsonSerializerFailureReason.LOOP_LIMIT_EXCEEDED;
END_METHOD

METHOD _serializeStatus : BOOL
VAR_IN_OUT
	v: SJsonValue;
END_VAR
VAR_INPUT
	pStatus: POINTER TO FB_Status;
END_VAR
VAR_OUTPUT
	failureReason: E_ProtoJsonSerializerFailureReason;
END_VAR
VAR
	_obj: SJsonValue;
	_member: SJsonValue;
END_VAR
_serializeStatus := FALSE;
failureReason := E_ProtoJsonSerializerFailureReason.NA;
IF v = 0 THEN
	failureReason := E_ProtoJsonSerializerFailureReason.JSON_VALUE_INVALID;
	RETURN;
END_IF
IF pStatus = 0 THEN
	failureReason := E_ProtoJsonSerializerFailureReason.VALUE_POINTER_NULL;
	RETURN;
END_IF

_obj := THIS^.parser.AddObjectMember(v, 'status');
IF _obj = 0 THEN
	failureReason := E_ProtoJsonSerializerFailureReason.JSON_OPERATION_FAILURE;
	RETURN;
END_IF
IF pStatus^.message <> 0 AND_THEN NOT THIS^.serializeStringValue(_obj, ADR('message'), pStatus^.message, failureReason=>failureReason) THEN
	RETURN;
END_IF
IF pStatus^.code <> E_StatusCode.STATUS_CODE_UNSET THEN
	_member := THIS^.parser.AddUintMember(_obj, 'code', TO_UDINT(pStatus^.code));
	IF _member = 0 THEN
		failureReason := E_ProtoJsonSerializerFailureReason.JSON_OPERATION_FAILURE;
		RETURN;
	END_IF
END_IF
_serializeStatus := failureReason = E_ProtoJsonSerializerFailureReason.NA;
END_METHOD

(* Appends one Span object to the JSON array v. The span is only read. *)
METHOD serializeSpan : BOOL
VAR_IN_OUT
	v: SJsonValue;
END_VAR
VAR_INPUT
	pSpan: POINTER TO FB_Span;
END_VAR
VAR_OUTPUT
	failureReason: E_ProtoJsonSerializerFailureReason;
END_VAR
VAR
	_obj: SJsonValue;
	_member: SJsonValue;
	_parentSpanId: STRING(16);
END_VAR
serializeSpan := FALSE;
failureReason := E_ProtoJsonSerializerFailureReason.NA;
IF v = 0 THEN
	failureReason := E_ProtoJsonSerializerFailureReason.JSON_VALUE_INVALID;
	RETURN;
END_IF
IF pSpan = 0 THEN
	failureReason := E_ProtoJsonSerializerFailureReason.SPAN_POINTER_NULL;
	RETURN;
END_IF

_obj := THIS^.parser.PushbackJsonValue(v, '{}');
IF _obj = 0 THEN
	failureReason := E_ProtoJsonSerializerFailureReason.JSON_OPERATION_FAILURE;
	RETURN;
END_IF

// identity; a root span has no parentSpanId
IF pSpan^.traceId <> 0 AND_THEN NOT THIS^.serializeTraceIdValue(_obj, pSpan^.traceId, failureReason=>failureReason) THEN RETURN; END_IF
IF pSpan^.spanId <> 0 AND_THEN NOT THIS^.serializeSpanIdValue(_obj, pSpan^.spanId, failureReason=>failureReason) THEN RETURN; END_IF
IF pSpan^.traceState <> 0 AND_THEN NOT THIS^._serializeTraceState(_obj, pSpan^.traceState, failureReason=>failureReason) THEN RETURN; END_IF
IF pSpan^.parentSpanId <> 0 THEN
	IF NOT THIS^._serializeBytes(
		ADR(pSpan^.parentSpanId^.bytes),
		SIZEOF(pSpan^.parentSpanId^.bytes),
		ADR(_parentSpanId),
		SIZEOF(_parentSpanId),
		E_BytesEncoding.hex,
		failureReason=>failureReason
	) THEN
		RETURN;
	END_IF
	_member := THIS^.parser.AddStringMember(_obj, 'parentSpanId', _parentSpanId);
	IF _member = 0 THEN failureReason := E_ProtoJsonSerializerFailureReason.JSON_OPERATION_FAILURE; RETURN; END_IF
END_IF
IF pSpan^.flags <> 0 AND_THEN NOT THIS^.serializeUint32Value(_obj, ADR('flags'), pSpan^.flags, failureReason=>failureReason) THEN RETURN; END_IF

// description and timing; OTLP/JSON writes enums as numbers and 64-bit integers as strings
IF pSpan^.name <> 0 AND_THEN NOT THIS^.serializeStringValue(_obj, ADR('name'), pSpan^.name, failureReason=>failureReason) THEN RETURN; END_IF
_member := THIS^.parser.AddUintMember(_obj, 'kind', TO_UDINT(pSpan^.kind));
IF _member = 0 THEN failureReason := E_ProtoJsonSerializerFailureReason.JSON_OPERATION_FAILURE; RETURN; END_IF
IF NOT THIS^.serializeUint64Value(_obj, ADR('startTimeUnixNano'), pSpan^.startTimestamp, failureReason=>failureReason) THEN RETURN; END_IF
IF NOT THIS^.serializeUint64Value(_obj, ADR('endTimeUnixNano'), pSpan^.endTimestamp, failureReason=>failureReason) THEN RETURN; END_IF

IF pSpan^.attributes.count > 0 AND_THEN NOT THIS^.serializeKeyValues(_obj, ADR('attributes'), ADR(pSpan^.attributes), failureReason=>failureReason) THEN RETURN; END_IF
IF pSpan^.attributes.droppedCount > 0 AND_THEN NOT THIS^.serializeUint32Value(
	_obj,
	ADR('droppedAttributesCount'),
	pSpan^.attributes.droppedCount,
	failureReason=>failureReason
) THEN
	RETURN;
END_IF
IF pSpan^.links.count > 0 AND_THEN NOT THIS^._serializeLinks(_obj, pSpan^.links, failureReason=>failureReason) THEN RETURN; END_IF
IF pSpan^.links.droppedCount > 0 AND_THEN NOT THIS^.serializeUint32Value(
	_obj,
	ADR('droppedLinksCount'),
	pSpan^.links.droppedCount,
	failureReason=>failureReason
) THEN
	RETURN;
END_IF
IF pSpan^.status <> 0 AND_THEN NOT THIS^._serializeStatus(_obj, pSpan^.status, failureReason=>failureReason) THEN RETURN; END_IF
serializeSpan := failureReason = E_ProtoJsonSerializerFailureReason.NA;
END_METHOD

METHOD startNewResource : BOOL
VAR_IN_OUT
	v: SJsonValue;
	resource: FB_Resource;
END_VAR
VAR_OUTPUT
	scopeSpans: SJsonValue;
	failureReason: E_ProtoJsonSerializerFailureReason;
END_VAR
VAR
	_resourceObj: SJsonValue;
	_member: SJsonValue;
END_VAR
startNewResource := FALSE;
scopeSpans := 0;
failureReason := E_ProtoJsonSerializerFailureReason.NA;
IF v = 0 THEN
	failureReason := E_ProtoJsonSerializerFailureReason.JSON_VALUE_INVALID;
	RETURN;
END_IF

_resourceObj := THIS^.parser.PushbackJsonValue(v, '{}');
IF _resourceObj = 0 THEN
	failureReason := E_ProtoJsonSerializerFailureReason.JSON_OPERATION_FAILURE;
	RETURN;
END_IF
IF NOT THIS^._injectResource(_resourceObj, resource, failureReason=>failureReason) THEN
	RETURN;
END_IF
IF resource.schemaUrl <> '' THEN
	_member := THIS^.parser.AddStringMember(_resourceObj, 'schemaUrl', resource.schemaUrl);
	IF _member = 0 THEN
		failureReason := E_ProtoJsonSerializerFailureReason.JSON_OPERATION_FAILURE;
		RETURN;
	END_IF
END_IF
scopeSpans := THIS^.parser.AddArrayMember(_resourceObj, 'scopeSpans', 0);
IF scopeSpans = 0 THEN
	failureReason := E_ProtoJsonSerializerFailureReason.JSON_OPERATION_FAILURE;
	RETURN;
END_IF

startNewResource := failureReason = E_ProtoJsonSerializerFailureReason.NA;
END_METHOD

METHOD startNewScope : BOOL
VAR_IN_OUT
	v: SJsonValue;
	scope: FB_InstrumentationScope;
END_VAR
VAR_OUTPUT
	serializedSpans: SJsonValue;
	failureReason: E_ProtoJsonSerializerFailureReason;
END_VAR
VAR
	_scopeObj: SJsonValue;
	_member: SJsonValue;
END_VAR
startNewScope := FALSE;
serializedSpans := 0;
failureReason := E_ProtoJsonSerializerFailureReason.NA;
IF v = 0 THEN
	failureReason := E_ProtoJsonSerializerFailureReason.JSON_VALUE_INVALID;
	RETURN;
END_IF

_scopeObj := THIS^.parser.PushbackJsonValue(v, '{}');
IF _scopeObj = 0 THEN
	failureReason := E_ProtoJsonSerializerFailureReason.JSON_OPERATION_FAILURE;
	RETURN;
END_IF
IF NOT THIS^._injectInstrumentationScope(_scopeObj, scope, failureReason=>failureReason) THEN
	RETURN;
END_IF
IF scope.schemaUrl <> '' THEN
	_member := THIS^.parser.AddStringMember(_scopeObj, 'schemaUrl', scope.schemaUrl);
	IF _member = 0 THEN
		failureReason := E_ProtoJsonSerializerFailureReason.JSON_OPERATION_FAILURE;
		RETURN;
	END_IF
END_IF
serializedSpans := THIS^.parser.AddArrayMember(_scopeObj, 'spans', 0);
IF serializedSpans = 0 THEN
	failureReason := E_ProtoJsonSerializerFailureReason.JSON_OPERATION_FAILURE;
	RETURN;
END_IF

startNewScope := failureReason = E_ProtoJsonSerializerFailureReason.NA;
END_METHOD

(*
	Writes one ResourceSpans group led by pSpan, which the caller has popped and owns. Every
	queued span of the same resource is popped and written, grouped by scope in first-seen
	order. Spans of other resources are rotated, so they keep their arrival order. pSpan is
	0 on success; on failure it holds any span still owned, for the caller to release.
*)
METHOD serializeResourceSpans : BOOL
VAR_IN_OUT
	v: SJsonValue;
	spans: FB_SpanQueue;
	pSpan: POINTER TO FB_Span;
END_VAR
VAR_OUTPUT
	failureReason: E_ProtoJsonSerializerFailureReason;
END_VAR
VAR
	_resourceId: UDINT;
	_scopeSpans: SJsonValue;
	_pHead: POINTER TO FB_Span;
	_scopeLimit: UDINT;
	_spansToScan: UDINT;
	_scopeIdx: UDINT;
	_scanIdx: UDINT;
	_queueFailureReason: E_SpanQueueFailureReason;
END_VAR
serializeResourceSpans := FALSE;
failureReason := E_ProtoJsonSerializerFailureReason.NA;
IF v = 0 THEN
	failureReason := E_ProtoJsonSerializerFailureReason.JSON_VALUE_INVALID;
	RETURN;
END_IF
IF pSpan = 0 THEN
	failureReason := E_ProtoJsonSerializerFailureReason.SPAN_POINTER_NULL;
	RETURN;
END_IF

_resourceId := pSpan^.resource.id;
IF NOT THIS^.startNewResource(
	v:=v,
	resource:=pSpan^.resource,
	scopeSpans=>_scopeSpans,
	failureReason=>failureReason
) THEN
	RETURN;
END_IF

// One scope per pass. Each pass writes at least the leading span, so count + 1 passes suffice.
_scopeLimit := spans.count + 1;
FOR _scopeIdx := 1 TO _scopeLimit DO
	IF NOT THIS^.serializeScopeSpans(
		v:=_scopeSpans,
		spans:=spans,
		pSpan:=pSpan,
		resourceId:=_resourceId,
		failureReason=>failureReason
	) THEN
		RETURN;
	END_IF

	// Pop the first span of another scope of this resource. Rotating every other span
	// preserves arrival order for later resource groups.
	_spansToScan := spans.count;
	FOR _scanIdx := 1 TO _spansToScan DO
		spans.reset();
		_pHead := spans.next();
		IF _pHead = 0 THEN
			failureReason := E_ProtoJsonSerializerFailureReason.SPAN_COLLECTION_INCONSISTENT;
			RETURN;
		END_IF
		IF pSpan = 0 AND_THEN _pHead^.resource.id = _resourceId THEN
			IF NOT spans.pop(pValue:=pSpan, failureReason=>_queueFailureReason) THEN
				failureReason := E_ProtoJsonSerializerFailureReason.QUEUE_POP_FAILURE;
				RETURN;
			END_IF
			IF pSpan = 0 THEN
				failureReason := E_ProtoJsonSerializerFailureReason.SPAN_COLLECTION_INCONSISTENT;
				RETURN;
			END_IF
		ELSIF NOT spans.rotate(failureReason=>_queueFailureReason) THEN
			failureReason := E_ProtoJsonSerializerFailureReason.QUEUE_ROTATE_FAILURE;
			RETURN;
		END_IF
	END_FOR

	IF pSpan = 0 THEN
		serializeResourceSpans := failureReason = E_ProtoJsonSerializerFailureReason.NA;
		RETURN;
	END_IF
END_FOR

failureReason := E_ProtoJsonSerializerFailureReason.LOOP_LIMIT_EXCEEDED;
END_METHOD

(*
	Writes one ScopeSpans group led by pSpan, which the caller has popped and owns. Every
	queued span with the same resource and scope is popped and written in queue order;
	other spans are rotated. Each span is released once written, so pSpan is 0 on success.
	On failure it holds any span still owned, for the caller to release.
*)
METHOD serializeScopeSpans : BOOL
VAR_IN_OUT
	v: SJsonValue;
	spans: FB_SpanQueue;
	pSpan: POINTER TO FB_Span;
END_VAR
VAR_INPUT
	resourceId: UDINT;
END_VAR
VAR_OUTPUT
	failureReason: E_ProtoJsonSerializerFailureReason;
END_VAR
VAR
	_scopeName: T_MaxString;
	_serializedSpans: SJsonValue;
	_pHead: POINTER TO FB_Span;
	_spansToScan: UDINT;
	_scanIdx: UDINT;
	_queueFailureReason: E_SpanQueueFailureReason;
END_VAR
serializeScopeSpans := FALSE;
failureReason := E_ProtoJsonSerializerFailureReason.NA;
IF v = 0 THEN
	failureReason := E_ProtoJsonSerializerFailureReason.JSON_VALUE_INVALID;
	RETURN;
END_IF
IF pSpan = 0 THEN
	failureReason := E_ProtoJsonSerializerFailureReason.SPAN_POINTER_NULL;
	RETURN;
END_IF
IF pSpan^.resource.id <> resourceId THEN
	failureReason := E_ProtoJsonSerializerFailureReason.SPAN_COLLECTION_INCONSISTENT;
	RETURN;
END_IF

_scopeName := pSpan^.scope.name;
IF NOT THIS^.startNewScope(
	v:=v,
	scope:=pSpan^.scope,
	serializedSpans=>_serializedSpans,
	failureReason=>failureReason
) THEN
	RETURN;
END_IF

IF NOT THIS^.serializeSpan(_serializedSpans, pSpan, failureReason=>failureReason) THEN
	RETURN;
END_IF
pSpan^.delete(pSelf:=pSpan);

// Consume and release every remaining span in this resource/scope group.
_spansToScan := spans.count;
FOR _scanIdx := 1 TO _spansToScan DO
	spans.reset();
	_pHead := spans.next();
	IF _pHead = 0 THEN
		failureReason := E_ProtoJsonSerializerFailureReason.SPAN_COLLECTION_INCONSISTENT;
		RETURN;
	END_IF

	IF _pHead^.resource.id = resourceId AND_THEN _pHead^.scope.name = _scopeName THEN
		IF NOT spans.pop(pValue:=pSpan, failureReason=>_queueFailureReason) THEN
			failureReason := E_ProtoJsonSerializerFailureReason.QUEUE_POP_FAILURE;
			RETURN;
		END_IF
		IF pSpan = 0 THEN
			failureReason := E_ProtoJsonSerializerFailureReason.SPAN_COLLECTION_INCONSISTENT;
			RETURN;
		END_IF
		IF NOT THIS^.serializeSpan(_serializedSpans, pSpan, failureReason=>failureReason) THEN
			RETURN;
		END_IF
		pSpan^.delete(pSelf:=pSpan);
	ELSIF NOT spans.rotate(failureReason=>_queueFailureReason) THEN
		failureReason := E_ProtoJsonSerializerFailureReason.QUEUE_ROTATE_FAILURE;
		RETURN;
	END_IF
END_FOR

serializeScopeSpans := failureReason = E_ProtoJsonSerializerFailureReason.NA;
END_METHOD

(*
	Writes a TracesData document for every span in the queue to jsonValue. Spans are grouped
	by resource and then by instrumentation scope, so each resource and scope is written once.
	Groups keep first-seen order, and spans keep queue order within a group.

	Takes ownership of all queued spans and drains the queue. Written spans are released as
	they are written, and any left over are released on failure, so the queue is empty
	whatever the result. Grouping rotates the queue once per group, so the work is bounded
	by count squared.
*)
METHOD serializeTracesData : BOOL
VAR_IN_OUT
	spans: FB_SpanQueue;
END_VAR
VAR_OUTPUT
	failureReason: E_ProtoJsonSerializerFailureReason;
END_VAR
VAR
	_count: UDINT;
	_pSpan: POINTER TO FB_Span;
	_resourceSpans: SJsonValue;
	_resourceIdx: UDINT;
	_queueFailureReason: E_SpanQueueFailureReason;
END_VAR
serializeTracesData := FALSE;
failureReason := E_ProtoJsonSerializerFailureReason.NA;

_count := spans.count;
IF _count > TcOtlp_GVL.MAX_LOOP_COUNT THEN
	spans.free();
	failureReason := E_ProtoJsonSerializerFailureReason.LOOP_LIMIT_EXCEEDED;
	RETURN;
END_IF

// start a new document whose root is an object holding the resourceSpans array
THIS^.jsonValue := THIS^.parser.NewDocument();
IF THIS^.jsonValue = 0 THEN
	spans.free();
	failureReason := E_ProtoJsonSerializerFailureReason.JSON_OPERATION_FAILURE;
	RETURN;
END_IF
THIS^.jsonValue := THIS^.parser.SetObject(THIS^.jsonValue);
IF THIS^.jsonValue = 0 THEN
	spans.free();
	failureReason := E_ProtoJsonSerializerFailureReason.JSON_OPERATION_FAILURE;
	RETURN;
END_IF
_resourceSpans := THIS^.parser.AddArrayMember(THIS^.jsonValue, 'resourceSpans', 0);
IF _resourceSpans = 0 THEN
	spans.free();
	failureReason := E_ProtoJsonSerializerFailureReason.JSON_OPERATION_FAILURE;
	RETURN;
END_IF

// each resource group pops at least its leading span, so _count passes always suffice
_pSpan := 0;
FOR _resourceIdx := 1 TO _count DO
	IF spans.count = 0 THEN
		EXIT;
	END_IF
	IF NOT spans.pop(pValue:=_pSpan, failureReason=>_queueFailureReason) THEN
		failureReason := E_ProtoJsonSerializerFailureReason.QUEUE_POP_FAILURE;
		EXIT;
	END_IF
	IF _pSpan = 0 THEN
		failureReason := E_ProtoJsonSerializerFailureReason.SPAN_COLLECTION_INCONSISTENT;
		EXIT;
	END_IF
	IF NOT THIS^.serializeResourceSpans(
		v:=_resourceSpans,
		spans:=spans,
		pSpan:=_pSpan,
		failureReason=>failureReason
	) THEN
		EXIT;
	END_IF
END_FOR

// release a span a failed group still holds
IF _pSpan <> 0 THEN
	_pSpan^.delete(pSelf:=_pSpan);
END_IF
IF failureReason = E_ProtoJsonSerializerFailureReason.NA AND spans.count > 0 THEN
	failureReason := E_ProtoJsonSerializerFailureReason.SPAN_COLLECTION_INCONSISTENT;
END_IF

spans.free();
serializeTracesData := failureReason = E_ProtoJsonSerializerFailureReason.NA;
END_METHOD

(*
	Writes a trace state as the traceState string member of v. OTLP carries the canonical W3C
	header as one string, which may be longer than T_MaxString.
*)
METHOD _serializeTraceState : BOOL
VAR_IN_OUT
	v: SJsonValue;
END_VAR
VAR_INPUT
	pTraceState: POINTER TO FB_TraceState;
END_VAR
VAR_OUTPUT
	failureReason: E_ProtoJsonSerializerFailureReason;
END_VAR
VAR
	_pText: POINTER TO STRING;
	_member: SJsonValue;
END_VAR
_serializeTraceState := FALSE;
failureReason := E_ProtoJsonSerializerFailureReason.NA;
IF v = 0 THEN failureReason := E_ProtoJsonSerializerFailureReason.JSON_VALUE_INVALID; RETURN; END_IF
IF pTraceState = 0 THEN failureReason := E_ProtoJsonSerializerFailureReason.VALUE_POINTER_NULL; RETURN; END_IF
_pText := pTraceState^.pString;
IF _pText = 0 THEN failureReason := E_ProtoJsonSerializerFailureReason.STRING_POINTER_NULL; RETURN; END_IF
_member := THIS^.parser.AddStringMember(v, 'traceState', _pText^);
IF _member = 0 THEN failureReason := E_ProtoJsonSerializerFailureReason.JSON_OPERATION_FAILURE; RETURN; END_IF
_serializeTraceState := TRUE;
END_METHOD

END_FUNCTION_BLOCK

// ---- OTEL/TRACING/PROCESSORS/FUNCTION_BLOCKS/FB_SpanProcessor_Batch.TcPOU
(*
	Keeps ended spans until they can be exported together. onEnd enriches the span and pushes a
	clone onto a bounded queue; nothing is exported during onEnd. tick advances the exporter and
	then, when the exporter is idle, hands it the oldest maxExportBatchSize spans once
	scheduledDelayMillis has passed since the queue became non-empty, or at once when a full
	batch is waiting. Spans that end in the same scan, or while the exporter is busy, therefore
	stay queued and go out in a later batch.
	When the queue holds maxQueueSize spans the oldest is dropped for the newest. droppedCount
	counts those spans and the spans that could not be cloned or queued.
	Pass 0 as the exporter to drop every span.
*)
FUNCTION_BLOCK FB_SpanProcessor_Batch EXTENDS FB_SpanProcessor_Base
VAR_OUTPUT
	scheduledDelayMillis: UDINT := 1000;  // maximum delay before queued spans are exported
	maxExportBatchSize: UDINT := 512;  // maximum spans handed to one export
	failureReason: E_SpanProcessorFailureReason;  // result of the last onEnd or export attempt
END_VAR
VAR
	_scheduleDelayTimer: TON;
	_spans: FB_SpanQueue(maxCount:=0);  // set again during THIS^.FB_Init
	_rejectedCount: UDINT;  // spans lost to clone or push failures
	_exporter: REFERENCE TO FB_SpanExporter_Base;
END_VAR

// no-op; override to change or add to the span before it is queued
METHOD enrich
VAR_IN_OUT
	span: FB_Span;
END_VAR
END_METHOD

(* Hands the oldest queued spans to an idle exporter when the delay has passed or a full batch waits. *)
METHOD exportIfNeeded
VAR
	_exportFailureReason: E_SpanExporterFailureReason;
END_VAR
IF THIS^.maxExportBatchSize = 0
	OR_ELSE NOT __ISVALIDREF(THIS^._exporter)
	OR_ELSE THIS^._exporter.isBusy()
	OR_ELSE THIS^._spans.count = 0 THEN
	RETURN;
END_IF

IF NOT THIS^._scheduleDelayTimer.Q
	AND_THEN THIS^._spans.count < THIS^.maxExportBatchSize THEN
	RETURN;
END_IF

// accepted spans move to the exporter; on failure they stay queued for the next attempt
IF THIS^._exporter.export(
	spans:=THIS^._spans,
	count:=THIS^.maxExportBatchSize,
	failureReason=>_exportFailureReason
) THEN
	THIS^._scheduleDelayTimer(IN:=FALSE, PT:=UDINT_TO_TIME(THIS^.scheduledDelayMillis));
	THIS^.failureReason := E_SpanProcessorFailureReason.NA;
ELSE
	THIS^.failureReason := E_SpanProcessorFailureReason.EXPORT_FAILURE;
END_IF
END_METHOD

METHOD FB_Exit : BOOL
VAR_INPUT
	bInCopyCode: BOOL;  // TRUE: the exit method is called in order to leave the instance which will be copied afterwards (online change).
END_VAR
IF NOT bInCopyCode THEN
	THIS^.free();
END_IF
END_METHOD

METHOD FB_Init : BOOL
VAR_INPUT
	bInitRetains: BOOL;  // TRUE: the retain variables are initialized (reset warm / reset cold)
	bInCopyCode: BOOL;  // TRUE: the instance will be copied to the copy code afterward (online change)
	maxQueueSize: UDINT := 2048;  // held to TcOtlp_GVL.MAX_LOOP_COUNT; zero means that limit
	scheduledDelayMillis: UDINT := 1000;  // maximum delay before queued spans are exported
	maxExportBatchSize: UDINT := 512;  // maximum spans handed to one export; zero never exports
	exporter: REFERENCE TO FB_SpanExporter_Base;  // borrowed and must outlive the processor; 0 drops every span
END_VAR
THIS^._spans.FB_Init(FALSE, FALSE, maxQueueSize);
THIS^.scheduledDelayMillis := scheduledDelayMillis;
THIS^.maxExportBatchSize := maxExportBatchSize;
IF __ISVALIDREF(exporter) THEN
	THIS^._exporter REF= exporter;
ELSE
	THIS^._exporter REF= 0;
END_IF
END_METHOD

(* Releases every queued span and restarts the schedule delay. *)
METHOD free
THIS^._spans.free();
THIS^._scheduleDelayTimer(IN:=FALSE, PT:=UDINT_TO_TIME(THIS^.scheduledDelayMillis));
END_METHOD

(*
	Enriches the borrowed span, then pushes a clone onto the queue. A full queue drops its
	oldest span to make room.
*)
METHOD onEnd
VAR_INPUT
	span: REFERENCE TO FB_Span;
END_VAR
VAR
	_pClone: POINTER TO FB_Span;
	_cloneFailureReason: E_SpanCloneFailureReason;
	_queueFailureReason: E_SpanQueueFailureReason;
END_VAR
IF NOT __ISVALIDREF(span) OR_ELSE NOT __ISVALIDREF(THIS^._exporter) THEN
	RETURN;
END_IF

THIS^.enrich(span);

IF NOT span.cloneTo(pDest:=_pClone, failureReason=>_cloneFailureReason) THEN
	IF _pClone <> 0 THEN _pClone^.delete(pSelf:=_pClone); END_IF
	THIS^._rejectedCount := THIS^._rejectedCount + 1;
	THIS^.failureReason := E_SpanProcessorFailureReason.SPAN_CLONE_FAILURE;
	RETURN;
END_IF

IF NOT THIS^._spans.push(pValue:=_pClone, failureReason=>_queueFailureReason) THEN
	_pClone^.delete(pSelf:=_pClone);
	THIS^._rejectedCount := THIS^._rejectedCount + 1;
	THIS^.failureReason := E_SpanProcessorFailureReason.QUEUE_PUSH_FAILURE;
	RETURN;
END_IF

THIS^.failureReason := E_SpanProcessorFailureReason.NA;
END_METHOD

(* Advances the exporter, then exports a batch if one is due. Called once per provider tick. *)
METHOD tick
VAR
	_exportFailureReason: E_SpanExporterFailureReason;
END_VAR
THIS^._scheduleDelayTimer(
	IN:=THIS^._spans.count > 0,
	PT:=UDINT_TO_TIME(THIS^.scheduledDelayMillis)
);

IF __ISVALIDREF(THIS^._exporter) THEN
	THIS^._exporter.tick(failureReason=>_exportFailureReason);
	THIS^.exportIfNeeded();
END_IF
END_METHOD

(* Spans lost so far: evicted from a full queue, or not cloned or queued. *)
PROPERTY droppedCount : UDINT
GET
droppedCount := THIS^._spans.droppedCount + THIS^._rejectedCount;
END_GET
END_PROPERTY

(* Spans waiting for export. *)
PROPERTY queuedCount : UDINT
GET
queuedCount := THIS^._spans.count;
END_GET
END_PROPERTY

END_FUNCTION_BLOCK

// ---- OTEL/TRACING/PROCESSORS/FUNCTION_BLOCKS/FB_SpanProcessor_Base.TcPOU
(*
	Contract for span processors. FB_TracerProvider stages processors each scan, then its tick
	passes every ended span to onEnd of each staged processor and releases the span once they
	have all returned. The span is borrowed: a processor that keeps it past onEnd must clone it.
*)
FUNCTION_BLOCK ABSTRACT FB_SpanProcessor_Base

(* Extension point that may change the span before it is exported. *)
METHOD ABSTRACT enrich
VAR_IN_OUT
	span: FB_Span;
END_VAR
END_METHOD

METHOD ABSTRACT free
END_METHOD

(* Called once for each ended span. The span is borrowed and released after the call. *)
METHOD ABSTRACT onEnd
VAR_INPUT
	span: REFERENCE TO FB_Span;
END_VAR
END_METHOD

PROPERTY pSelf : POINTER TO FB_SpanProcessor_Base
GET
pSelf := THIS;
END_GET
END_PROPERTY

(* Called once per provider tick, after the ended spans have been handed out. *)
METHOD ABSTRACT tick
END_METHOD

END_FUNCTION_BLOCK

// ---- OTEL/TRACING/EXPORTING/FUNCTION_BLOCKS/FB_SpanExporter_Console.TcPOU
(*
	Writes one line per span to the TwinCAT ADS log at hint level, for development and
	commissioning. For example:
	  span "work" trace=0101...01 span=0202020202020202 parent=none kind=SPAN_KIND_INTERNAL status=STATUS_CODE_UNSET duration=500ns
	export writes the whole batch and releases it before returning, so the exporter is never
	busy and suits FB_SpanProcessor_Simple. Attributes, links, resource and scope are not
	written. Lines longer than 255 characters are truncated.
*)
FUNCTION_BLOCK FB_SpanExporter_Console EXTENDS FB_SpanExporter_Base

THIS^.tick(failureReason=>THIS^._callFailureReason);

(* Lower-case hex of count bytes; at most 64 bytes are written. *)
METHOD _hex : T_MaxString
VAR_INPUT
	pBytes: POINTER TO BYTE;
	count: UDINT;
END_VAR
VAR CONSTANT
	MAX_BYTES: UDINT := 64;
END_VAR
VAR
	_i: UDINT;
END_VAR
_hex := '';
IF pBytes = 0 THEN
	RETURN;
END_IF

FOR _i := 1 TO MIN(count, MAX_BYTES) DO
	_hex := CONCAT(_hex, BYTE_TO_HEXSTR(in:=pBytes[_i - 1], iPrecision:=2, bLoCase:=TRUE));
END_FOR
END_METHOD

(* Accepts the batch, writes one line per span and releases the batch. *)
METHOD export : BOOL
VAR_IN_OUT
	spans: FB_SpanQueue;
END_VAR
VAR_INPUT
	count: UDINT;
END_VAR
VAR_OUTPUT
	failureReason: E_SpanExporterFailureReason;
END_VAR
VAR
	_idx: UDINT;
	_pSpan: POINTER TO FB_Span;
END_VAR
export := SUPER^.export(
	spans:=spans,
	count:=count,
	failureReason=>failureReason
);
IF NOT export THEN
	RETURN;
END_IF

THIS^._spans.reset();
FOR _idx := 1 TO TcOtlp_GVL.MAX_LOOP_COUNT DO
	_pSpan := THIS^._spans.next();
	IF _pSpan = 0 THEN
		EXIT;
	END_IF
	ADSLOGSTR(msgCtrlMask:=ADSLOG_MSGTYPE_HINT, msgFmtStr:='%s', strArg:=THIS^.format(_pSpan^));
END_FOR

THIS^.free();
END_METHOD

(* Builds the log line for one span. Missing members are written as empty, none or unset. *)
METHOD format : T_MaxString
VAR_INPUT
	span: REFERENCE TO FB_Span;
END_VAR
VAR
	_name: T_MaxString;
	_traceId: T_MaxString;
	_spanId: T_MaxString;
	_parent: T_MaxString := 'none';
	_status: E_StatusCode := E_StatusCode.STATUS_CODE_UNSET;
	_duration: ULINT;
END_VAR
format := '';
IF NOT __ISVALIDREF(span) THEN
	RETURN;
END_IF

IF span.name <> 0 AND_THEN span.name^.pString <> 0 THEN
	_name := span.name^.pString^;
END_IF
IF span.traceId <> 0 THEN
	_traceId := THIS^._hex(pBytes:=ADR(span.traceId^.bytes), count:=SIZEOF(span.traceId^.bytes));
END_IF
IF span.spanId <> 0 THEN
	_spanId := THIS^._hex(pBytes:=ADR(span.spanId^.bytes), count:=SIZEOF(span.spanId^.bytes));
END_IF
IF span.parentSpanId <> 0 THEN
	_parent := THIS^._hex(pBytes:=ADR(span.parentSpanId^.bytes), count:=SIZEOF(span.parentSpanId^.bytes));
END_IF
IF span.status <> 0 THEN
	_status := span.status^.code;
END_IF
IF span.endTimestamp > span.startTimestamp THEN
	_duration := span.endTimestamp - span.startTimestamp;
END_IF

format := CONCAT('span "', _name);
format := CONCAT(format, '" trace=');
format := CONCAT(format, _traceId);
format := CONCAT(format, ' span=');
format := CONCAT(format, _spanId);
format := CONCAT(format, ' parent=');
format := CONCAT(format, _parent);
format := CONCAT(format, ' kind=');
format := CONCAT(format, TO_STRING(span.kind));
format := CONCAT(format, ' status=');
format := CONCAT(format, TO_STRING(_status));
format := CONCAT(format, ' duration=');
format := CONCAT(format, ULINT_TO_STRING(_duration));
format := CONCAT(format, 'ns');
END_METHOD

METHOD isBusy : BOOL
isBusy := FALSE;
END_METHOD

METHOD tick : BOOL
VAR_OUTPUT
	failureReason: E_SpanExporterFailureReason;
END_VAR
failureReason := E_SpanExporterFailureReason.NA;
tick := TRUE;
END_METHOD

END_FUNCTION_BLOCK

// ---- OTEL/TRACING/EXPORTING/FUNCTION_BLOCKS/FB_SpanExporter_HTTP.TcPOU
(*
	Posts each accepted batch as one OTLP/HTTP ProtoJSON TracesData request to an OTLP
	collector, for example 'http://192.168.1.10:4318/v1/traces'. Call the instance, or tick,
	every scan: the exporter is busy from export until currentState reaches done or error.
	The batch is released at either end, and an error is reported by tick until the next
	batch is accepted. A response outside 2xx is an error; nothing is retried.
*)
FUNCTION_BLOCK FB_SpanExporter_HTTP EXTENDS FB_SpanExporter_Base
VAR_OUTPUT
	currentState: E_HttpExporterState;
	statusCode: UINT;  // the HTTP status code received for the last completed request
END_VAR

VAR
	_execute: BOOL;
	_urlParsed: BOOL;
	_endpoint: ST_HttpEndpoint;
	_len: UDINT;
	_execRTrig: R_TRIG;
	_pString: POINTER TO STRING;
	_jsonVal: SJsonValue;
	_computedState: E_HttpExporterState;
	_failureReason: E_SpanExporterFailureReason;
	_serializationFailureReason: E_ProtoJsonSerializerFailureReason;
	_serializer: FB_SpanProtoJsonSerializer;
	_client: FB_IotHttpClient;
	_request: FB_IotHttpRequest;
	_header: FB_IotHttpHeaderFieldMap;
END_VAR

THIS^.tick(failureReason=>THIS^._callFailureReason);

METHOD export: BOOL
VAR_IN_OUT
	spans: FB_SpanQueue;
END_VAR
VAR_INPUT
	count: UDINT;
END_VAR
VAR_OUTPUT
	failureReason: E_SpanExporterFailureReason;
END_VAR
// a finished exporter accepts the next batch at once
IF THIS^.currentState = E_HttpExporterState.done OR THIS^.currentState = E_HttpExporterState.error THEN
	THIS^.currentState := E_HttpExporterState.idle;
	THIS^._computedState := E_HttpExporterState.idle;
END_IF
export := SUPER^.export(
	spans:=spans,
	count:=count,
	failureReason=>failureReason
);
IF export THEN
	THIS^._failureReason := E_SpanExporterFailureReason.NA;
	THIS^._serializationFailureReason := E_ProtoJsonSerializerFailureReason.NA;
END_IF
END_METHOD

(*
	Releases a payload buffer that is still in flight. The FB_IotHttpRequest reading it is
	destroyed with this instance, so nothing uses the buffer afterwards. TwinCAT then
	runs FB_SpanExporter_Base.FB_Exit, which releases the accepted spans.
*)
METHOD FB_Exit : BOOL
VAR_INPUT
	bInCopyCode: BOOL;  // TRUE: the instance is being copied during an online change
END_VAR
// during an online change the copy keeps the buffer, so it must not be released here
IF NOT bInCopyCode AND _pString <> 0 THEN
	__DELETE(_pString);
	_pString := 0;
END_IF
END_METHOD

METHOD FB_Init: BOOL
VAR_INPUT
	bInitRetains: BOOL; // TRUE: the retain variables are initialized (reset warm / reset cold)
	bInCopyCode: BOOL;  // TRUE: the instance will be copied to the copy code afterward (online change)
	url: T_MaxString;  // full endpoint URL, e.g. 'http://192.168.1.10:4318/v1/traces'
	bNoServerCertCheck: BOOL := FALSE;  // allow HTTPS connections to servers with self-signed certificates
END_VAR
THIS^.currentState := E_HttpExporterState.idle;
THIS^._computedState := E_HttpExporterState.idle;

THIS^._urlParsed := F_ParseHttpUrl(url:=url, endpoint=>THIS^._endpoint);

THIS^._client.sHostName := THIS^._endpoint.host;
THIS^._client.nHostPort := THIS^._endpoint.port;
THIS^._client.bKeepAlive := TRUE;
THIS^._client.tConnectionTimeout := T#10S;
IF THIS^._endpoint.useTls THEN
	THIS^._client.stTLS.bNoServerCertCheck := bNoServerCertCheck;
END_IF

THIS^._request.sContentType := 'application/json';
END_METHOD

METHOD isBusy : BOOL
isBusy := THIS^._exportActive;
END_METHOD

METHOD tick : BOOL
VAR_OUTPUT
	failureReason: E_SpanExporterFailureReason;
END_VAR
tick := TRUE;
failureReason := E_SpanExporterFailureReason.NA;

_execute := THIS^._exportActive;
_execRTrig(CLK := _execute AND_THEN THIS^._spans.count > 0);

CASE currentState OF
	E_HttpExporterState.idle:
		IF _execRTrig.Q THEN
			_failureReason := E_SpanExporterFailureReason.NA;
			_serializationFailureReason := E_ProtoJsonSerializerFailureReason.NA;
			IF NOT THIS^._urlParsed THEN
				_failureReason := E_SpanExporterFailureReason.HTTP_URL_PARSE_FAILURE;
				_computedState := E_HttpExporterState.error;
			ELSE
				_computedState := E_HttpExporterState.serializing;
			END_IF
		END_IF

	E_HttpExporterState.serializing:
		// the serializer drains the batch; buffer the TracesData document as the payload
		IF NOT _serializer.serializeTracesData(
			spans:=THIS^._spans,
			failureReason=>_serializationFailureReason
		) THEN
			_failureReason := E_SpanExporterFailureReason.SERIALIZATION_FAILURE;
			_computedState := E_HttpExporterState.error;
		ELSE
			_jsonVal := _serializer.jsonValue;
			IF _jsonVal = 0 OR_ELSE NOT _serializer.parser.IsObject(_jsonVal) THEN
				_failureReason := E_SpanExporterFailureReason.SERIALIZATION_FAILURE;
				_computedState := E_HttpExporterState.error;
			ELSE
				_len := _serializer.parser.GetJsonLength(_jsonVal);  // includes the null terminating character
				IF _len = 0 THEN
					_failureReason := E_SpanExporterFailureReason.SERIALIZATION_FAILURE;
					_computedState := E_HttpExporterState.error;
				ELSE
					_pString := __NEW(BYTE, _len);
					IF _pString = 0 THEN
						_failureReason := E_SpanExporterFailureReason.BUFFER_ALLOCATION_FAILURE;
						_computedState := E_HttpExporterState.error;
					ELSE
						_serializer.parser.CopyJson(_jsonVal, _pString^, _len);
						_computedState := E_HttpExporterState.sending;
					END_IF
				END_IF
			END_IF
		END_IF

	E_HttpExporterState.sending:
		IF NOT _request.bBusy THEN
			IF _request.SendRequest(
				sUri := THIS^._endpoint.path,
				fbClient := THIS^._client,
				eRequestType := ETcIotHttpRequestType.HTTP_POST,
				pContent := _pString,
				nContentSize := _len - 1,
				fbHeader := THIS^._header
			) THEN
				_computedState := E_HttpExporterState.waiting;
			ELSE
				IF _pString <> 0 THEN __DELETE(_pString); _pString := 0; END_IF
				_failureReason := E_SpanExporterFailureReason.HTTP_REQUEST_FAILURE;
				_computedState := E_HttpExporterState.error;
			END_IF
		END_IF

	E_HttpExporterState.waiting:
		IF NOT _request.bBusy THEN
			_computedState := E_HttpExporterState.processing;
		END_IF

	E_HttpExporterState.processing:
		IF _request.bError THEN
			IF _pString <> 0 THEN __DELETE(_pString); _pString := 0; END_IF
			_failureReason := E_SpanExporterFailureReason.HTTP_REQUEST_FAILURE;
			_computedState := E_HttpExporterState.error;
		ELSE
			statusCode := _request.nStatusCode;
			IF statusCode < 200 OR_ELSE statusCode >= 300 THEN
				IF _pString <> 0 THEN __DELETE(_pString); _pString := 0; END_IF
				_failureReason := E_SpanExporterFailureReason.HTTP_STATUS_FAILURE;
				_computedState := E_HttpExporterState.error;
			ELSE
				IF _pString <> 0 THEN __DELETE(_pString); _pString := 0; END_IF
				_computedState := E_HttpExporterState.done;
			END_IF
		END_IF

	E_HttpExporterState.done:
		IF NOT _execute THEN
			_computedState := E_HttpExporterState.idle;
		END_IF

	E_HttpExporterState.error:
		// keep the failure until export accepts a new batch
END_CASE

currentState := _computedState;

IF currentState = E_HttpExporterState.done
	OR_ELSE currentState = E_HttpExporterState.error THEN
	THIS^.free();
END_IF

THIS^._client.Execute();

IF currentState = E_HttpExporterState.error THEN
	tick := FALSE;
	failureReason := _failureReason;
END_IF
END_METHOD

END_FUNCTION_BLOCK

// ---- OTEL/TRACING/PROPAGATION/TraceContextPropagator.TcPOU
(*
	Decodes W3C Trace Context carriers into span contexts, and encodes span contexts into them.
	Propagation is the caller's job: the application owns the carrier, the transport and the span
	it starts, and this program only converts between a context and an ST_TraceContextCarrier.
	It knows nothing about how a carrier travels, so each transport (ADS, OPC UA, HTTP) is a
	separate block that moves the carrier and calls inject or extract. See "Trace Context
	Propagation" in the docs.
*)
PROGRAM TraceContextPropagator
VAR CONSTANT
	TRACEPARENT_LENGTH: UDINT := 55;  // version 00, and the fields every version starts with: 2 + 1 + 32 + 1 + 16 + 1 + 2
	TRACE_ID_OFFSET: UDINT := 3;
	SPAN_ID_OFFSET: UDINT := 36;
	FLAGS_OFFSET: UDINT := 53;
	DELIMITER: BYTE := 16#2D;  // '-'
	MAX_TRACESTATE_LENGTH: UDINT := 512;  // the W3C floor for propagating a tracestate; the size of ST_TraceContextCarrier.tracestate
END_VAR

(*
	Parses a W3C traceparent and optional tracestate into a new remote span context. The caller
	owns pDest, which must be 0, and releases it once with delete. Nothing is allocated until the
	traceparent is known to be good, and on failure pDest stays 0: the caller should then start
	its span without the context, because a mangled header must not stop a process.
	An all-zero trace id or span id is the encoding of "absent" and is rejected. Version ff is
	invalid. Version 00 is exactly 55 characters; a future version may be longer, and is read as
	its first 55 characters when the flags are followed by '-'. The headers are taken by
	reference at their full length, so an overlong traceparent is seen and rejected, and the
	tracestate is never cut mid-entry. W3C asks for at least 512 tracestate characters to be
	kept and allows only whole entries to be dropped, so every entry is kept here; a carrier of
	limited size uses TraceStateFactory.truncate when the context is sent on. An invalid
	tracestate is dropped without failing the extraction. The context is marked remote. The
	default sampler follows its sampled bit for a span that takes it as a parent, and ignores it
	for a span that only links to it.
*)
METHOD extract : BOOL
VAR_IN_OUT
	pDest: POINTER TO FB_SpanContext;
END_VAR
VAR_IN_OUT CONSTANT
	traceparent: STRING;  // any length: pass carrier.traceparent, or a longer header as received
	tracestate: STRING;  // any length; '' when the header is absent
END_VAR
VAR_OUTPUT
	failureReason: E_PropagationFailureReason;
END_VAR
VAR
	_p: POINTER TO BYTE;
	_length: UDINT;
	_allZero: BOOL;
	_version: BYTE;
	_flags: BYTE;
	_traceId: FB_TraceId;
	_spanId: FB_SpanId;
	_pTraceState: POINTER TO FB_TraceState;
END_VAR
extract := FALSE;
failureReason := E_PropagationFailureReason.NA;

IF pDest <> 0 THEN
	failureReason := E_PropagationFailureReason.DESTINATION_ALREADY_ASSIGNED;
	RETURN;
END_IF

// measured with LEN2, because LEN stops at 255 characters
_p := ADR(traceparent);
_length := TO_UDINT(LEN2(_p));

IF _length = 0 THEN
	failureReason := E_PropagationFailureReason.TRACEPARENT_EMPTY;
	RETURN;
END_IF

IF _length < TRACEPARENT_LENGTH THEN
	failureReason := E_PropagationFailureReason.TRACEPARENT_LENGTH_INVALID;
	RETURN;
END_IF

// every field sits at a fixed offset, so validation is a bounded decode of 27 bytes
IF NOT _decodeHex(pText:=_p, nBytes:=1, pBytes:=ADR(_version)) OR_ELSE _version = 16#FF THEN
	failureReason := E_PropagationFailureReason.VERSION_INVALID;
	RETURN;
END_IF

// version 00 has no room for more fields
IF _version = 0 AND _length > TRACEPARENT_LENGTH THEN
	failureReason := E_PropagationFailureReason.TRACEPARENT_LENGTH_INVALID;
	RETURN;
END_IF

// a future version may add fields after the flags, each introduced by '-'
IF _p[TRACE_ID_OFFSET - 1] <> DELIMITER
	OR _p[SPAN_ID_OFFSET - 1] <> DELIMITER
	OR _p[FLAGS_OFFSET - 1] <> DELIMITER
	OR (_length > TRACEPARENT_LENGTH AND_THEN _p[TRACEPARENT_LENGTH] <> DELIMITER)
THEN
	failureReason := E_PropagationFailureReason.DELIMITER_INVALID;
	RETURN;
END_IF

IF NOT _decodeHex(
		pText:=_p + TRACE_ID_OFFSET,
		nBytes:=SIZEOF(_traceId.bytes),
		pBytes:=ADR(_traceId.bytes),
		allZero=>_allZero)
	OR _allZero
THEN
	failureReason := E_PropagationFailureReason.TRACE_ID_INVALID;
	RETURN;
END_IF

IF NOT _decodeHex(
		pText:=_p + SPAN_ID_OFFSET,
		nBytes:=SIZEOF(_spanId.bytes),
		pBytes:=ADR(_spanId.bytes),
		allZero=>_allZero)
	OR _allZero
THEN
	failureReason := E_PropagationFailureReason.SPAN_ID_INVALID;
	RETURN;
END_IF

IF NOT _decodeHex(pText:=_p + FLAGS_OFFSET, nBytes:=1, pBytes:=ADR(_flags)) THEN
	failureReason := E_PropagationFailureReason.TRACE_FLAGS_INVALID;
	RETURN;
END_IF

// the traceparent is good; an invalid tracestate leaves _pTraceState at 0 and is dropped
TraceStateFactory.parse(pDest:=_pTraceState, pHeader:=ADR(tracestate));

IF NOT ContextFactory.buildContext(
	pDest:=pDest,
	pTraceId:=ADR(_traceId),
	pSpanId:=ADR(_spanId),
	pTraceState:=_pTraceState,
	traceFlags:=TO_UDINT(_flags)
		OR TO_UDINT(E_SpanFlags.SPAN_FLAGS_CONTEXT_HAS_IS_REMOTE_MASK)
		OR TO_UDINT(E_SpanFlags.SPAN_FLAGS_CONTEXT_IS_REMOTE_MASK))
THEN
	failureReason := E_PropagationFailureReason.MEMORY_ALLOCATION_FAILURE;
END_IF

// the context holds its own copy of the trace state
IF _pTraceState <> 0 THEN _pTraceState^.delete(pSelf:=_pTraceState); END_IF

extract := failureReason = E_PropagationFailureReason.NA;
END_METHOD

(*
	Decodes nBytes bytes from the 2 * nBytes hex characters at pText into pBytes. W3C allows
	only lowercase hex, so any other character fails. allZero reports whether every decoded
	byte is 0. nBytes comes from the fixed traceparent fields, so it is at most 16.
*)
METHOD _decodeHex : BOOL
VAR_INPUT
	pText: POINTER TO BYTE;
	nBytes: UDINT;
	pBytes: POINTER TO BYTE;
END_VAR
VAR_OUTPUT
	allZero: BOOL;
END_VAR
VAR
	_i: UDINT;
	_high: BYTE;
	_low: BYTE;
END_VAR
_decodeHex := FALSE;
allZero := TRUE;

IF pText = 0 OR pBytes = 0 OR nBytes = 0 THEN
	RETURN;
END_IF

FOR _i := 0 TO nBytes - 1 DO
	_high := _hexValue(pText[2 * _i]);
	_low := _hexValue(pText[2 * _i + 1]);
	IF _high > 15 OR _low > 15 THEN
		RETURN;
	END_IF
	pBytes[_i] := SHL(_high, 4) OR _low;
	allZero := allZero AND pBytes[_i] = 0;
END_FOR

_decodeHex := TRUE;
END_METHOD

(* Returns the value of one lowercase hex digit, or 16#FF when c is not one. *)
METHOD _hexValue : BYTE
VAR_INPUT
	c: BYTE;
END_VAR
IF c >= 16#30 AND c <= 16#39 THEN  // '0'..'9'
	_hexValue := c - 16#30;
ELSIF c >= 16#61 AND c <= 16#66 THEN  // 'a'..'f'
	_hexValue := c - 16#61 + 10;
ELSE
	_hexValue := 16#FF;
END_IF
END_METHOD

(*
	Writes a span context into a carrier, for an outbound call. The context is borrowed and not
	changed. The traceparent is version 00 with the low 8 bits of the trace
	flags, which are the W3C trace flags; the OTLP remote bits are not propagated. A trace state
	longer than MAX_TRACESTATE_LENGTH is shortened with TraceStateFactory.truncate, which drops
	whole entries as W3C requires, and a context without one writes ''. On failure both headers
	are left empty, so a caller never sends half a carrier.
*)
METHOD inject : BOOL
VAR_INPUT
	pContext: POINTER TO FB_SpanContext;
END_VAR
VAR_IN_OUT
	carrier: ST_TraceContextCarrier;
END_VAR
VAR_OUTPUT
	failureReason: E_PropagationFailureReason;
END_VAR
VAR
	_p: POINTER TO BYTE;
	_flags: BYTE;
	_pSource: POINTER TO FB_TraceState;
	_pShort: POINTER TO FB_TraceState;
END_VAR
inject := FALSE;
failureReason := E_PropagationFailureReason.NA;
carrier.traceparent := '';
carrier.tracestate := '';

IF pContext = 0 THEN
	failureReason := E_PropagationFailureReason.CONTEXT_POINTER_NULL;
	RETURN;
END_IF

IF NOT pContext^.isValid() THEN
	failureReason := E_PropagationFailureReason.CONTEXT_INVALID;
	RETURN;
END_IF

// the trace state first: it is the only step that can fail after validation
_pSource := pContext^.traceState;
IF _pSource <> 0 AND_THEN _pSource^.length > MAX_TRACESTATE_LENGTH THEN
	// the context's trace state was validated when it was parsed, so only allocation can fail
	IF NOT TraceStateFactory.truncate(pDest:=_pShort, pSrc:=_pSource, maxLength:=MAX_TRACESTATE_LENGTH) THEN
		failureReason := E_PropagationFailureReason.MEMORY_ALLOCATION_FAILURE;
		RETURN;
	END_IF
	_pSource := _pShort;  // 0 when no entry fits, which writes ''
END_IF
IF _pSource <> 0 THEN
	MEMCPY(destAddr:=ADR(carrier.tracestate), srcAddr:=_pSource^.pString, n:=_pSource^.length);
	_p := ADR(carrier.tracestate);
	_p[_pSource^.length] := 0;
END_IF
IF _pShort <> 0 THEN _pShort^.delete(pSelf:=_pShort); END_IF

// every field sits at a fixed offset: 00-<trace id>-<span id>-<flags>
_p := ADR(carrier.traceparent);
_p[0] := 16#30;  // '0'
_p[1] := 16#30;
_p[TRACE_ID_OFFSET - 1] := DELIMITER;
_encodeHex(pBytes:=ADR(pContext^.traceId.bytes), nBytes:=SIZEOF(pContext^.traceId.bytes), pText:=_p + TRACE_ID_OFFSET);
_p[SPAN_ID_OFFSET - 1] := DELIMITER;
_encodeHex(pBytes:=ADR(pContext^.spanId.bytes), nBytes:=SIZEOF(pContext^.spanId.bytes), pText:=_p + SPAN_ID_OFFSET);
_p[FLAGS_OFFSET - 1] := DELIMITER;
_flags := TO_BYTE(pContext^.traceFlags AND 16#FF);
_encodeHex(pBytes:=ADR(_flags), nBytes:=1, pText:=_p + FLAGS_OFFSET);
_p[TRACEPARENT_LENGTH] := 0;

inject := TRUE;
END_METHOD

(*
	Writes nBytes bytes from pBytes as 2 * nBytes lowercase hex characters at pText, the only
	case W3C allows. nBytes comes from the fixed traceparent fields, so it is at most 16.
*)
METHOD _encodeHex
VAR_INPUT
	pBytes: POINTER TO BYTE;
	nBytes: UDINT;
	pText: POINTER TO BYTE;
END_VAR
VAR
	_i: UDINT;
END_VAR
IF pBytes = 0 OR pText = 0 OR nBytes = 0 THEN
	RETURN;
END_IF

FOR _i := 0 TO nBytes - 1 DO
	pText[2 * _i] := _hexDigit(SHR(pBytes[_i], 4));
	pText[2 * _i + 1] := _hexDigit(pBytes[_i] AND 16#0F);
END_FOR
END_METHOD

(* Returns the lowercase hex character for a value from 0 to 15. *)
METHOD _hexDigit : BYTE
VAR_INPUT
	value: BYTE;
END_VAR
IF value < 10 THEN
	_hexDigit := 16#30 + value;  // '0'..'9'
ELSE
	_hexDigit := 16#57 + value;  // 'a'..'f': 16#61 - 10
END_IF
END_METHOD

END_PROGRAM

// ---- OTEL/TRACING/SAMPLING/FUNCTION_BLOCKS/FB_Sampler_AlwaysOn.TcPOU
(*
	Samples every span, as the OpenTelemetry AlwaysOn sampler does, even the child of a parent
	that was not sampled.
*)
FUNCTION_BLOCK FB_Sampler_AlwaysOn EXTENDS FB_Sampler

METHOD onStart
VAR_INPUT
	span: REFERENCE TO FB_Span;
END_VAR
span.setSampled(TRUE);
END_METHOD

END_FUNCTION_BLOCK

// ---- OTEL/TRACING/SAMPLING/FUNCTION_BLOCKS/FB_Sampler_ErrorsOnly.TcPOU
(*
	Keeps only the sampled spans that end with STATUS_CODE_ERROR, so a controller exports the
	operations that failed and nothing else. The start decision is the default one, so a failed
	span whose parent was not sampled is still dropped.
*)
FUNCTION_BLOCK FB_Sampler_ErrorsOnly EXTENDS FB_Sampler

(* Drops a span that has no status or ended with an OK status. *)
METHOD onEnd
VAR_INPUT
	span: REFERENCE TO FB_Span;
END_VAR
IF span.status = 0 OR_ELSE span.status^.code <> E_StatusCode.STATUS_CODE_ERROR THEN
	span.setSampled(FALSE);
END_IF
END_METHOD

END_FUNCTION_BLOCK

// ---- OTEL/TRACING/ID_GENERATION/FUNCTION_BLOCKS/FB_IdGenerator.TcPOU
FUNCTION_BLOCK FB_IdGenerator EXTENDS FB_IdGenerator_Base
VAR CONSTANT
	GUID_BYTES: UDINT := 16;  // one guid, which is also the width of a trace id
END_VAR
VAR
	_creator: Tc2_System.FB_CreateGUID;
	_pBuffer: POINTER TO BYTE;
	_bufferLen: UDINT;
	_head: POINTER TO BYTE;
	_tail: POINTER TO BYTE;
	_count: UDINT;  // unread bytes, starting at _head
	_headRoom: UDINT;  // bytes from _head to the end of the ring, never zero
	_tailRoom: UDINT;  // bytes from _tail to the end of the ring, never zero
	_inFlight: UDINT;  // bytes the refill in flight will write at _tail, 0 when none is out
	_edgeHeld: BOOL;  // bExecute has been high for a cycle, so bBusy describes this request
END_VAR
VAR_OUTPUT
	errorId: UDINT;  // last ADS error reported by the guid service, 0 when healthy
END_VAR

(* Cuts nBytes off the head of the ring into pDest, which must have room for them.
   pDest is borrowed for the duration of the call and never taken. *)
METHOD _take : BOOL
VAR_INPUT
	pDest: POINTER TO BYTE;
	nBytes: UDINT;
END_VAR
VAR_OUTPUT
	failureReason: E_IdGenFailureReason;
END_VAR
VAR
	_first: UDINT;  // bytes of the draw that lie ahead of _head, before the ring wraps
END_VAR
_take := FALSE;
failureReason := E_IdGenFailureReason.NA;

IF NOT THIS^.configValid THEN
	failureReason := E_IdGenFailureReason.INVALID_CONFIGUATION;
	RETURN;
END_IF

// a draw wider than the ring itself can never be served, however long the caller waits,
// so it is reported as the configuration mistake it is rather than as an empty ring
IF (pDest = 0) OR_ELSE (nBytes = 0) OR_ELSE (nBytes > THIS^._bufferLen) THEN
	failureReason := E_IdGenFailureReason.INVALID_CONFIGUATION;
	RETURN;
END_IF

// nothing is written until the draw is known to be servable, which is what leaves the
// caller's identifier untouched on failure
IF THIS^._count < nBytes THEN
	failureReason := E_IdGenFailureReason.NO_IDENTIFIERS_AVAILABLE;
	RETURN;
END_IF

// a draw may straddle the wrap, so it is stitched from the bytes ahead of _head and, once
// those run out, the bytes at the start of the ring. A refill is never stitched this way,
// which is why only this side of the ring has to know about the seam.
_first := THIS^._headRoom;
IF _first > nBytes THEN
	_first := nBytes;
END_IF

MEMCPY(pDest, THIS^._head, _first);
IF _first < nBytes THEN
	MEMCPY(pDest + _first, THIS^._pBuffer, nBytes - _first);
END_IF

// Advance the read point over what was taken. _tail is deliberately left alone: that is
// what keeps the destination of a refill in flight from moving out from under it.
IF _first < THIS^._headRoom THEN
	THIS^._head := THIS^._head + nBytes;
	THIS^._headRoom := THIS^._headRoom - nBytes;
ELSE
	// the draw reached the end of the ring, so reading resumes at its start
	THIS^._head := THIS^._pBuffer + (nBytes - _first);
	THIS^._headRoom := THIS^._bufferLen - (nBytes - _first);
END_IF

THIS^._count := THIS^._count - nBytes;
_take := TRUE;
END_METHOD

PROPERTY configValid : BOOL
GET
configValid := THIS^._pBuffer <> 0;
END_GET
END_PROPERTY

//FB_Exit must be implemented explicitly. If there is an implementation, then the
//method is called before the controller removes the code of the function block instance
//(implicit call). The return value is not evaluated.
METHOD FB_Exit: BOOL
VAR_INPUT
    bInCopyCode: BOOL;  // TRUE: the exit method is called in order to leave the instance which will be copied afterwards (online change).  
END_VAR
IF NOT bInCopyCode THEN
	THIS^.free();
END_IF
END_METHOD

//FB_Init is always available implicitly and it is used primarily for initialization.
//The return value is not evaluated. For a specific influence, you can also declare the
//methods explicitly and provide additional code there with the standard initialization
//code. You can evaluate the return value.
METHOD FB_Init: BOOL
VAR_INPUT
    bInitRetains: BOOL; // TRUE: the retain variables are initialized (reset warm / reset cold)
    bInCopyCode: BOOL;  // TRUE: the instance will be copied to the copy code afterward (online change)
	nTraceIds: UDINT;
	nSpanIds: UDINT;
END_VAR
IF (NOT bInCopyCode) AND nTraceIds > 0 AND nSpanIds > 0 THEN
	THIS^._bufferLen := ((nTraceIds*16) + (nSpanIds*8));

	// the ring grows up to a whole number of guids. The guid service writes nothing smaller
	// than one, so a remainder shorter than a guid could never be filled, and because the
	// fill point cannot skip over a hole the ring would strand at the wrap.
	IF (THIS^._bufferLen MOD GUID_BYTES) <> 0 THEN
		THIS^._bufferLen := THIS^._bufferLen + (GUID_BYTES - (THIS^._bufferLen MOD GUID_BYTES));
	END_IF

	THIS^._pBuffer := __NEW(BYTE, THIS^._bufferLen);
	THIS^._head := THIS^._pBuffer;
	THIS^._tail := THIS^._pBuffer;
	THIS^._headRoom := THIS^._bufferLen;
	THIS^._tailRoom := THIS^._bufferLen;
END_IF
END_METHOD

(*
	Releases the ring and resets every cursor into it. Safe to call more than once.
	A refill still in flight is abandoned: tick stops calling the guid service once
	configValid is FALSE, so the service is never handed the released buffer again.
*)
METHOD free
IF THIS^._pBuffer <> 0 THEN
	__DELETE(THIS^._pBuffer);
	THIS^._pBuffer := 0;
END_IF
THIS^._bufferLen := 0;
THIS^._head := 0;
THIS^._tail := 0;
THIS^._count := 0;
THIS^._headRoom := 0;
THIS^._tailRoom := 0;
THIS^._inFlight := 0;
THIS^._edgeHeld := FALSE;
END_METHOD

METHOD generateSpanId : BOOL
VAR_IN_OUT
	spanId: FB_SpanId;
END_VAR
VAR_OUTPUT
	failureReason: E_IdGenFailureReason;
END_VAR
// the identifier states its own width, so the draw is eight bytes without anyone here
// having to name the number
generateSpanId := THIS^._take(
	pDest:=ADR(spanId.bytes),
	nBytes:=TO_UDINT(SIZEOF(spanId.bytes)),
	failureReason=>failureReason
);
END_METHOD

METHOD generateTraceId : BOOL
VAR_IN_OUT
	traceId: FB_TraceId;
END_VAR
VAR_OUTPUT
	failureReason: E_IdGenFailureReason;
END_VAR
// sixteen bytes, taken from the same ring as a span id, because the two identifiers are
// only different widths of the same random bytes
generateTraceId := THIS^._take(
	pDest:=ADR(traceId.bytes),
	nBytes:=TO_UDINT(SIZEOF(traceId.bytes)),
	failureReason=>failureReason
);
END_METHOD

(* Drives the refill request that keeps the ring populated. *)
METHOD tick : BOOL
VAR_OUTPUT
	failureReason: E_IdGenFailureReason;
END_VAR
VAR
	_room: UDINT;  // bytes the next refill may claim, before it is cut to whole guids
END_VAR
tick := FALSE;
failureReason := E_IdGenFailureReason.NA;

IF NOT THIS^.configValid THEN
	failureReason := E_IdGenFailureReason.INVALID_CONFIGUATION;
	RETURN;
END_IF

// The service writes one contiguous region, so a refill starts at _tail and stops at the
// end of the ring. Free space on the far side of the wrap is left to the refill after this
// one, because filling that side first would leave a hole at _tail and a ring has no way
// to describe a hole.
//
// The service is only ever handed the region _inFlight claims, which is what proves the
// region lies inside the allocation, and its length is remembered rather than recomputed
// because takes move _head while the request is out. A take never moves _tail, so the
// destination cannot shift out from under a request in flight.
THIS^._creator(
	bExecute := (THIS^._inFlight > 0),
	pGuidBuffer := THIS^._tail,
	nGuidBufferSize := THIS^._inFlight
);

IF THIS^._inFlight = 0 THEN
	// Nothing is out, so claim the room from _tail to the end of the ring, bounded by the
	// free space when that runs out first and cut to whole guids. bExecute is only raised by
	// the call above on the next cycle, which leaves the service a low cycle to see the edge.
	_room := THIS^._bufferLen - THIS^._count;
	IF _room > THIS^._tailRoom THEN
		_room := THIS^._tailRoom;
	END_IF
	THIS^._inFlight := (_room / GUID_BYTES) * GUID_BYTES;

ELSIF NOT THIS^._edgeHeld THEN
	// bBusy does not describe this request until the service has seen bExecute high
	THIS^._edgeHeld := TRUE;

ELSIF THIS^._creator.bError THEN
	// a failed request never advances _count, so the bytes it did not write are never
	// handed out as identifiers
	THIS^.errorId := THIS^._creator.nErrorId;
	THIS^._inFlight := 0;
	THIS^._edgeHeld := FALSE;
	failureReason := E_IdGenFailureReason.GUID_SERVICE_FAILED;
	RETURN;

ELSIF NOT THIS^._creator.bBusy THEN
	// the bytes are written, so publish them by advancing the fill point over them
	THIS^.errorId := 0;
	THIS^._count := THIS^._count + THIS^._inFlight;
	THIS^._tail := THIS^._tail + THIS^._inFlight;
	THIS^._tailRoom := THIS^._tailRoom - THIS^._inFlight;
	IF THIS^._tailRoom = 0 THEN
		THIS^._tail := THIS^._pBuffer;
		THIS^._tailRoom := THIS^._bufferLen;
	END_IF
	THIS^._inFlight := 0;
	THIS^._edgeHeld := FALSE;
END_IF

tick := TRUE;
END_METHOD

END_FUNCTION_BLOCK

// ---- OTEL/TRACING/ID_GENERATION/FUNCTION_BLOCKS/FB_IdGenerator_Base.TcPOU
(* Produces the trace and span identifiers that tracers attach to new spans.
   This is the only place in the tracing domain that creates identifier values;
   every other function block borrows or copies them.

   Implementations must never emit an all zero identifier, because an all zero
   identifier is the OTLP representation of "invalid/absent":
     - a trace id is 16 bytes and MUST NOT be all zeroes,
     - a span id is 8 bytes and MUST NOT be all zeroes.

   Generation is separated from span creation because it is not guaranteed to be
   constant time work. The owning provider calls `call` once per cycle to advance
   any bounded per cycle work; tracers only take finished identifiers. An
   implementation may therefore have nothing to hand out yet, in which case
   generation fails with NO_IDENTIFIERS_AVAILABLE instead of blocking the cycle. *)
FUNCTION_BLOCK ABSTRACT FB_IdGenerator_Base

(* Produces one valid, non zero span id into the caller owned spanId.
   Returns FALSE without modifying spanId on failure. *)
METHOD ABSTRACT generateSpanId : BOOL
VAR_IN_OUT
	spanId: FB_SpanId;
END_VAR
VAR_OUTPUT
	failureReason: E_IdGenFailureReason;
END_VAR
END_METHOD

(* Produces one valid, non zero trace id into the caller owned traceId.
   Returns FALSE without modifying traceId on failure. *)
METHOD ABSTRACT generateTraceId : BOOL
VAR_IN_OUT
	traceId: FB_TraceId;
END_VAR
VAR_OUTPUT
	failureReason: E_IdGenFailureReason;
END_VAR
END_METHOD

(* Advances any bounded per cycle generation work.
   Invoked by the owning provider, not by tracers.
   Returns FALSE and reports a failure reason when the generator cannot advance. *)
METHOD ABSTRACT tick : BOOL
VAR_OUTPUT
	failureReason: E_IdGenFailureReason;
END_VAR
END_METHOD

END_FUNCTION_BLOCK

// ---- OTEL/TRACING/PROCESSORS/FUNCTION_BLOCKS/FB_SpanProcessor_Simple.TcPOU
(*
	Handles each ended span as soon as the provider hands it over: enrich, then export.
	export clones the span and offers the clone to the exporter as a batch of one. The span is
	dropped when the exporter is busy or the clone fails, and nothing is kept between calls.
	Pass 0 as the exporter to drop every span, or override export to send spans somewhere
	else. Use FB_SpanExporter_Console to write spans to the ADS log.
*)
FUNCTION_BLOCK FB_SpanProcessor_Simple EXTENDS FB_SpanProcessor_Base
VAR
	_spans: FB_SpanQueue(maxCount:=1);
	_exporter: REFERENCE TO FB_SpanExporter_Base;
END_VAR

// no-op; override to change or add to the span before it is exported
METHOD enrich
VAR_IN_OUT
	span: FB_Span;
END_VAR
END_METHOD

(* Sends one ended span on. The span is borrowed for the duration of the call, so the
   exporter is given a clone, which it owns once it accepts it. *)
METHOD export
VAR_INPUT
	span: REFERENCE TO FB_Span;
END_VAR
VAR
	_pClone: POINTER TO FB_Span;
	_cloneFailureReason: E_SpanCloneFailureReason;
	_queueFailureReason: E_SpanQueueFailureReason;
	_exportFailureReason: E_SpanExporterFailureReason;
END_VAR
IF NOT __ISVALIDREF(THIS^._exporter) OR_ELSE THIS^._exporter.isBusy() THEN
	RETURN;
END_IF

IF span.cloneTo(pDest:=_pClone, failureReason=>_cloneFailureReason)
	AND_THEN THIS^._spans.push(pValue:=_pClone, failureReason=>_queueFailureReason) THEN
	THIS^._exporter.export(spans:=THIS^._spans, count:=1, failureReason=>_exportFailureReason);
END_IF

// whatever the exporter did not accept is dropped
THIS^._spans.free();
IF _pClone <> 0 THEN _pClone^.delete(pSelf:=_pClone); END_IF
END_METHOD

METHOD FB_Exit : BOOL
VAR_INPUT
	bInCopyCode: BOOL;  // TRUE: the exit method is called in order to leave the instance which will be copied afterwards (online change).
END_VAR
IF NOT bInCopyCode THEN
	THIS^.free();
END_IF
END_METHOD

// the simple processor keeps nothing between calls; this releases a span left by a failed hand-off
METHOD free
THIS^._spans.free();
END_METHOD

METHOD onEnd
VAR_INPUT
	span: REFERENCE TO FB_Span;
END_VAR
IF NOT __ISVALIDREF(span) THEN
	RETURN;
END_IF

THIS^.enrich(span);
THIS^.export(span);
END_METHOD

// advances the exporter's delivery once per provider tick
METHOD tick
VAR
	_exportFailureReason: E_SpanExporterFailureReason;
END_VAR
IF __ISVALIDREF(THIS^._exporter) THEN
	THIS^._exporter.tick(failureReason=>_exportFailureReason);
END_IF
END_METHOD

METHOD FB_Init : BOOL
VAR_INPUT
	bInitRetains: BOOL;  // TRUE: the retain variables are initialized (reset warm / reset cold)
	bInCopyCode: BOOL;  // TRUE: the instance will be copied to the copy code afterward (online change)
	exporter: REFERENCE TO FB_SpanExporter_Base;  // borrowed and must outlive the processor; 0 drops every span
END_VAR
IF __ISVALIDREF(exporter) THEN
	THIS^._exporter REF= exporter;
ELSE
	THIS^._exporter REF= 0;
END_IF
END_METHOD

END_FUNCTION_BLOCK

// ---- OTEL/TRACING/PROVIDER/FUNCTION_BLOCKS/FB_TracerProvider.TcPOU
(*
	Owns the ended spans of every tracer created from it and hands them to processors.
	Stage the processors every scan, then call tick once; tick passes each ended span to
	every staged processor, releases the span, and clears the staged list.
	The sampler decides which ended spans reach the processors; see onEnd.

	Example:
	provider.stageProcessor(consoleProcessor);
	// ... tracers start and end spans ...
	provider.tick(failureReason => reason);
*)
FUNCTION_BLOCK FB_TracerProvider
VAR
	_resource: REFERENCE TO FB_Resource;  // borrowed; the declaring scope owns its lifetime
	_idGenerator: REFERENCE TO FB_IdGenerator_Base;  // borrowed; the declaring scope owns its lifetime
	_sampler: REFERENCE TO FB_Sampler;  // borrowed; the declaring scope owns its lifetime
	_spans: FB_SpanQueue(TcOtlp_GVL.MAX_SPAN_RECORDS_PER_SCAN);  // ended spans waiting to be processed
	_head: POINTER TO ST_LinkedListNode;  // staged processors; the nodes are owned, the processors borrowed
	_failureReason: E_TracerProviderFailureReason;  // first staging failure since the last tick
END_VAR
VAR_OUTPUT
	stagedProcessorCount: UDINT;
END_VAR

(* Releases the staged-list nodes. The processors themselves are borrowed and untouched. *)
METHOD _freeProcessors
VAR
	_idx: UDINT;
	_node: POINTER TO ST_LinkedListNode;
END_VAR
FOR _idx := 0 TO TcOtlp_GVL.MAX_LOOP_COUNT DO
	IF THIS^._head = 0 THEN
		EXIT;
	END_IF
	_node := THIS^._head^.nxt;
	__DELETE(THIS^._head);
	THIS^._head := _node;
	// count down per node, so the count never claims nodes that are gone or hides ones that remain
	IF THIS^.stagedProcessorCount > 0 THEN
		THIS^.stagedProcessorCount := THIS^.stagedProcessorCount - 1;
	END_IF
END_FOR
END_METHOD

METHOD FB_Exit : BOOL
VAR_INPUT
	bInCopyCode: BOOL;  // TRUE: the exit method is called in order to leave the instance which will be copied afterwards (online change).
END_VAR
IF NOT bInCopyCode THEN
	THIS^._freeProcessors();
END_IF
END_METHOD

//FB_Init is always available implicitly and it is used primarily for initialization.
//The return value is not evaluated. For a specific influence, you can also declare the
//methods explicitly and provide additional code there with the standard initialization
//code. You can evaluate the return value.
METHOD FB_Init: BOOL
VAR_INPUT
    bInitRetains: BOOL; // TRUE: the retain variables are initialized (reset warm / reset cold)
    bInCopyCode: BOOL;  // TRUE: the instance will be copied to the copy code afterward (online change)
	resource: REFERENCE TO FB_Resource;
	idGenerator: REFERENCE TO FB_IdGenerator_Base;  // the source of identifiers for every tracer of this provider
	sampler: REFERENCE TO FB_Sampler;  // decides which spans are sampled; TcOtlp_GVL.defaultSampler is the OpenTelemetry default
END_VAR
THIS^._resource REF= resource;
THIS^._idGenerator REF= idGenerator;
THIS^._sampler REF= sampler;
END_METHOD

(*
	Takes ownership of an ended span and queues it for processing. On success pSpan is
	cleared; on failure it is left unchanged and still owned by the caller.
	A span that is not sampled is released instead, and that counts as success. The sampler's
	onEnd is asked only about spans that are still sampled, so it can drop a span but never
	keep one that its onStart dropped.
*)
METHOD onEnd : BOOL
VAR_IN_OUT
	pSpan: POINTER TO FB_Span;
END_VAR
VAR
	_pushFailureReason: E_SpanQueueFailureReason;
END_VAR
IF pSpan = 0 THEN
	RETURN;
END_IF

